screen "9" 800x480, template "Template_2"
   Button "Button_1" at 38,239 size 120x40; TextOff 'Carbamazepine'
      on Click: ActivateScreen("4_ORDER", 0); SetTag("Selected_URL", 'file:///C:/ASRS_Video/clip181.html')
      on Activate: SetTag("Selected_Medicine", 181)
      on Release: SetTag("ยา 181", 0)
      on Press: SetTag("ยา 181", 1)
   Button "Button_10" at 38,415 size 120x40; TextOff 'Pioglitazone'
      on Click: ActivateScreen("4_ORDER", 0); SetTag("Selected_URL", 'file:///C:/ASRS_Video/clip186.html')
      on Activate: SetTag("Selected_Medicine", 186)
      on Release: SetTag("ยา 186", 0)
      on Press: SetTag("ยา 186", 1)
   Button "Button_2" at 189,240 size 120x40; TextOff 'Levetiracetam'
      on Click: ActivateScreen("4_ORDER", 0); SetTag("Selected_URL", 'file:///C:/ASRS_Video/clip182.html')
      on Activate: SetTag("Selected_Medicine", 182)
      on Release: SetTag("ยา 182", 0)
      on Press: SetTag("ยา 182", 1)
   Button "Button_3" at 190,415 size 120x40; TextOff 'Sitagliptin'
      on Click: ActivateScreen("4_ORDER", 0); SetTag("Selected_URL", 'file:///C:/ASRS_Video/clip187.html')
      on Activate: SetTag("Selected_Medicine", 187)
      on Release: SetTag("ยา 187", 0)
      on Press: SetTag("ยา 187", 1)
   Button "Button_4" at 340,240 size 120x40; TextOff 'Metformin'
      on Click: ActivateScreen("4_ORDER", 0); SetTag("Selected_URL", 'file:///C:/ASRS_Video/clip183.html')
      on Activate: SetTag("Selected_Medicine", 183)
      on Release: SetTag("ยา 183", 0)
      on Press: SetTag("ยา 183", 1)
   Button "Button_5" at 340,416 size 120x40; TextOff 'Insulin regular'
      on Click: ActivateScreen("4_ORDER", 0); SetTag("Selected_URL", 'file:///C:/ASRS_Video/clip188.html')
      on Activate: SetTag("Selected_Medicine", 188)
      on Release: SetTag("ยา 188", 0)
      on Press: SetTag("ยา 188", 1)
   Button "Button_6" at 492,416 size 120x40; TextOff 'Insulin NPH'
      on Click: ActivateScreen("4_ORDER", 0); SetTag("Selected_URL", 'file:///C:/ASRS_Video/clip189.html')
      on Activate: SetTag("Selected_Medicine", 189)
      on Release: SetTag("ยา 189", 0)
      on Press: SetTag("ยา 189", 1)
   Button "Button_7" at 492,240 size 120x40; TextOff 'Glibenclamide'
      on Click: ActivateScreen("4_ORDER", 0); SetTag("Selected_URL", 'file:///C:/ASRS_Video/clip184.html')
      on Activate: SetTag("Selected_Medicine", 184)
      on Release: SetTag("ยา 184", 0)
      on Press: SetTag("ยา 184", 1)
   Button "Button_8" at 644,240 size 120x40; TextOff 'Gliclazide'
      on Click: ActivateScreen("4_ORDER", 0); SetTag("Selected_URL", 'file:///C:/ASRS_Video/clip185.html')
      on Activate: SetTag("Selected_Medicine", 185)
      on Release: SetTag("ยา 185", 0)
      on Press: SetTag("ยา 185", 1)
   Button "Button_11" at 645,416 size 120x40; TextOff 'Insulin glargine'
      on Click: ActivateScreen("4_ORDER", 0); SetTag("Selected_URL", 'file:///C:/ASRS_Video/clip190.html')
      on Activate: SetTag("Selected_Medicine", 190)
      on Release: SetTag("ยา 190", 0)
      on Press: SetTag("ยา 190", 1)
   Button "Button_12" at 24,16 size 94x40; TextOff 'Back'
      on Press: ActivateScreen("8", 0)
   Button "Button_9" at 688,16 size 96x40; TextOff 'Next'
      on Press: ActivateScreen("10", 0)
   GraphicView "Template_Graphic view_2" at 27,19 size 36x32; Picture "fast-backward"
   GraphicView "Template_Graphic view_1" at 693,20 size 36x32; Picture "play"
   GraphicView "Template_Graphic view_3" at 37,128 size 120x104; Picture "Picture181"
   GraphicView "Template_Graphic view_4" at 191,129 size 120x104; Picture "Picture182"
   GraphicView "Template_Graphic view_5" at 339,129 size 120x104; Picture "Picture183"
   GraphicView "Template_Graphic view_6" at 493,129 size 120x104; Picture "Picture184"
   GraphicView "Template_Graphic view_7" at 645,129 size 120x104; Picture "Picture185"
   GraphicView "Template_Graphic view_8" at 38,305 size 120x104; Picture "Picture186"
   GraphicView "Template_Graphic view_9" at 189,304 size 120x112; Picture "Picture187"
   GraphicView "Template_Graphic view_10" at 351,307 size 96x104; Picture "Picture188"
   GraphicView "Template_Graphic view_11" at 497,304 size 120x112; Picture "Picture189"
   GraphicView "Template_Graphic view_12" at 645,304 size 120x104; Picture "Picture190"
   TextField "Template_Text field_2" at 201,80 size 20x32; Text '9'

screen "10" 800x480, template "Template_2"
   Button "Button_1" at 38,239 size 120x40; TextOff 'Levothyroxine'
      on Click: ActivateScreen("4_ORDER", 0); SetTag("Selected_URL", 'file:///C:/ASRS_Video/clip191.html')
      on Activate: SetTag("Selected_Medicine", 191)
      on Release: SetTag("ยา 191", 0)
      on Press: SetTag("ยา 191", 1)
   Button "Button_10" at 38,415 size 120x40; TextOff 'Hydrocortisone'
      on Click: ActivateScreen("4_ORDER", 0); SetTag("Selected_URL", 'file:///C:/ASRS_Video/clip196.html')
      on Activate: SetTag("Selected_Medicine", 196)
      on Release: SetTag("ยา 196", 0)
      on Press: SetTag("ยา 196", 1)
   Button "Button_2" at 189,240 size 120x40; TextOff 'Propylthiouracil'
      on Click: ActivateScreen("4_ORDER", 0); SetTag("Selected_URL", 'file:///C:/ASRS_Video/clip192.html')
      on Activate: SetTag("Selected_Medicine", 192)
      on Release: SetTag("ยา 192", 0)
      on Press: SetTag("ยา 192", 1)
   Button "Button_3" at 190,415 size 120x40; TextOff 'Colchicine'
      on Click: ActivateScreen("4_ORDER", 0); SetTag("Selected_URL", 'file:///C:/ASRS_Video/clip197.html')
      on Activate: SetTag("Selected_Medicine", 197)
      on Release: SetTag("ยา 197", 0)
      on Press: SetTag("ยา 197", 1)
   Button "Button_4" at 340,240 size 120x40; TextOff 'Methimazole'
      on Click: ActivateScreen("4_ORDER", 0); SetTag("Selected_URL", 'file:///C:/ASRS_Video/clip193.html')
      on Activate: SetTag("Selected_Medicine", 193)
      on Release: SetTag("ยา 193", 0)
      on Press: SetTag("ยา 193", 1)
   Button "Button_5" at 340,416 size 120x40; TextOff 'Allopurinol'
      on Click: ActivateScreen("4_ORDER", 0); SetTag("Selected_URL", 'file:///C:/ASRS_Video/clip198.html')
      on Activate: SetTag("Selected_Medicine", 198)
      on Release: SetTag("ยา 198", 0)
      on Press: SetTag("ยา 198", 1)
   Button "Button_6" at 492,416 size 120x40; TextOff 'Febuxostat'
      on Click: ActivateScreen("4_ORDER", 0); SetTag("Selected_URL", 'file:///C:/ASRS_Video/clip199.html')
      on Activate: SetTag("Selected_Medicine", 199)
      on Release: SetTag("ยา 199", 0)
      on Press: SetTag("ยา 199", 1)
   Button "Button_7" at 492,240 size 120x40; TextOff 'Prednisolone'
      on Click: ActivateScreen("4_ORDER", 0); SetTag("Selected_URL", 'file:///C:/ASRS_Video/clip194.html')
      on Activate: SetTag("Selected_Medicine", 194)
      on Release: SetTag("ยา 194", 0)
      on Press: SetTag("ยา 194", 1)
   Button "Button_8" at 644,240 size 120x40; TextOff 'Dexamethasone'
      on Click: ActivateScreen("4_ORDER", 0); SetTag("Selected_URL", 'file:///C:/ASRS_Video/clip195.html')
      on Activate: SetTag("Selected_Medicine", 195)
      on Release: SetTag("ยา 195", 0)
      on Press: SetTag("ยา 195", 1)
   Button "Button_11" at 645,416 size 120x40; TextOff 'Calcium carbonate'
      on Click: ActivateScreen("4_ORDER", 0); SetTag("Selected_URL", 'file:///C:/ASRS_Video/clip200.html')
      on Activate: SetTag("Selected_Medicine", 200)
      on Release: SetTag("ยา 200", 0)
      on Press: SetTag("ยา 200", 1)
   Button "Button_12" at 24,16 size 94x40; TextOff 'Back'
      on Press: ActivateScreen("9", 0)
   Button "Button_9" at 688,16 size 96x40; TextOff 'Next'
      on Press: ActivateScreen("11", 0)
   GraphicView "Template_Graphic view_2" at 27,19 size 36x32; Picture "fast-backward"
   GraphicView "Template_Graphic view_1" at 693,20 size 36x32; Picture "play"
   GraphicView "Template_Graphic view_3" at 37,128 size 120x104; Picture "Picture191"
   GraphicView "Template_Graphic view_4" at 191,129 size 120x104; Picture "Picture192"
   GraphicView "Template_Graphic view_5" at 339,129 size 120x104; Picture "Picture193"
   GraphicView "Template_Graphic view_6" at 493,129 size 120x104; Picture "Picture194"
   GraphicView "Template_Graphic view_7" at 645,129 size 120x104; Picture "Picture195"
   GraphicView "Template_Graphic view_8" at 38,305 size 120x104; Picture "Picture196"
   GraphicView "Template_Graphic view_9" at 189,304 size 120x112; Picture "Picture197"
   GraphicView "Template_Graphic view_10" at 351,307 size 96x104; Picture "Picture198"
   GraphicView "Template_Graphic view_11" at 497,304 size 120x112; Picture "Picture199"
   GraphicView "Template_Graphic view_12" at 645,304 size 120x104; Picture "Picture200"
   TextField "Template_Text field_2" at 201,80 size 36x32; Text '10'

screen "11" 800x480, template "Template_2"
   Button "Button_1" at 38,239 size 120x40; TextOff 'Vitamin B complex'
      on Click: ActivateScreen("4_ORDER", 0); SetTag("Selected_URL", 'file:///C:/ASRS_Video/clip201.html')
      on Activate: SetTag("Selected_Medicine", 201)
      on Release: SetTag("ยา 201", 0)
      on Press: SetTag("ยา 201", 1)
   Button "Button_10" at 38,415 size 120x40; TextOff 'Potassium chloride'
      on Click: ActivateScreen("4_ORDER", 0); SetTag("Selected_URL", 'file:///C:/ASRS_Video/clip206.html')
      on Activate: SetTag("Selected_Medicine", 206)
      on Release: SetTag("ยา 206", 0)
      on Press: SetTag("ยา 206", 1)
   Button "Button_2" at 189,240 size 120x40; TextOff 'Vitamin C'
      on Click: ActivateScreen("4_ORDER", 0); SetTag("Selected_URL", 'file:///C:/ASRS_Video/clip202.html')
      on Activate: SetTag("Selected_Medicine", 202)
      on Release: SetTag("ยา 202", 0)
      on Press: SetTag("ยา 202", 1)
   Button "Button_3" at 190,415 size 120x40; TextOff 'Sodium bicarbonate'
      on Click: ActivateScreen("4_ORDER", 0); SetTag("Selected_URL", 'file:///C:/ASRS_Video/clip207.html')
      on Activate: SetTag("Selected_Medicine", 207)
      on Release: SetTag("ยา 207", 0)
      on Press: SetTag("ยา 207", 1)
   Button "Button_4" at 340,240 size 120x40; TextOff 'Ferrous fumarate'
      on Click: ActivateScreen("4_ORDER", 0); SetTag("Selected_URL", 'file:///C:/ASRS_Video/clip203.html')
      on Activate: SetTag("Selected_Medicine", 203)
      on Release: SetTag("ยา 203", 0)
      on Press: SetTag("ยา 203", 1)
   Button "Button_5" at 340,416 size 120x40; TextOff 'Calcium gluconate'
      on Click: ActivateScreen("4_ORDER", 0); SetTag("Selected_URL", 'file:///C:/ASRS_Video/clip208.html')
      on Activate: SetTag("Selected_Medicine", 208)
      on Release: SetTag("ยา 208", 0)
      on Press: SetTag("ยา 208", 1)
   Button "Button_6" at 492,416 size 120x40; TextOff 'Magnesium sulfate'
      on Click: ActivateScreen("4_ORDER", 0); SetTag("Selected_URL", 'file:///C:/ASRS_Video/clip209.html')
      on Activate: SetTag("Selected_Medicine", 209)
      on Release: SetTag("ยา 209", 0)
      on Press: SetTag("ยา 209", 1)
   Button "Button_7" at 492,240 size 120x40; TextOff 'Folic acid'
      on Click: ActivateScreen("4_ORDER", 0); SetTag("Selected_URL", 'file:///C:/ASRS_Video/clip204.html')
      on Activate: SetTag("Selected_Medicine", 204)
      on Release: SetTag("ยา 204", 0)
      on Press: SetTag("ยา 204", 1)
   Button "Button_8" at 644,240 size 120x40; TextOff 'Cyanocobalamin'
      on Click: ActivateScreen("4_ORDER", 0); SetTag("Selected_URL", 'file:///C:/ASRS_Video/clip205.html')
      on Activate: SetTag("Selected_Medicine", 205)
      on Release: SetTag("ยา 205", 0)
      on Press: SetTag("ยา 205", 1)
   Button "Button_11" at 645,416 size 120x40; TextOff 'Multivitamin'
      on Click: ActivateScreen("4_ORDER", 0); SetTag("Selected_URL", 'file:///C:/ASRS_Video/clip210.html')
      on Activate: SetTag("Selected_Medicine", 210)
      on Release: SetTag("ยา 210", 0)
      on Press: SetTag("ยา 210", 1)
   Button "Button_12" at 24,16 size 94x40; TextOff 'Back'
      on Press: ActivateScreen("10", 0)
   Button "Button_9" at 688,16 size 96x40; TextOff 'Next'
      on Press: ActivateScreen("12", 0)
   GraphicView "Template_Graphic view_2" at 27,19 size 36x32; Picture "fast-backward"
   GraphicView "Template_Graphic view_1" at 693,20 size 36x32; Picture "play"
   GraphicView "Template_Graphic view_3" at 37,128 size 120x104; Picture "Picture201"
   GraphicView "Template_Graphic view_4" at 191,129 size 120x104; Picture "Picture202"
   GraphicView "Template_Graphic view_5" at 339,129 size 120x104; Picture "Picture203"
   GraphicView "Template_Graphic view_6" at 493,129 size 120x104; Picture "Picture204"
   GraphicView "Template_Graphic view_7" at 645,129 size 120x104; Picture "Picture205"
   GraphicView "Template_Graphic view_8" at 38,305 size 120x104; Picture "Picture206"
   GraphicView "Template_Graphic view_9" at 189,304 size 120x112; Picture "Picture207"
   GraphicView "Template_Graphic view_10" at 351,307 size 96x104; Picture "Picture208"
   GraphicView "Template_Graphic view_11" at 497,304 size 120x112; Picture "Picture209"
   GraphicView "Template_Graphic view_12" at 645,304 size 120x104; Picture "Picture210"
   TextField "Template_Text field_2" at 201,80 size 36x32; Text '11'

screen "12" 800x480, template "Template_2"
   Button "Button_1" at 38,239 size 120x40; TextOff 'Oral rehydration salt'
      on Click: ActivateScreen("4_ORDER", 0); SetTag("Selected_URL", 'file:///C:/ASRS_Video/clip211.html')
      on Activate: SetTag("Selected_Medicine", 211)
      on Release: SetTag("ยา 211", 0)
      on Press: SetTag("ยา 211", 1)
   Button "Button_10" at 38,415 size 120x40; TextOff 'Piroxicam'
      on Click: ActivateScreen("4_ORDER", 0); SetTag("Selected_URL", 'file:///C:/ASRS_Video/clip216.html')
      on Activate: SetTag("Selected_Medicine", 216)
      on Release: SetTag("ยา 216", 0)
      on Press: SetTag("ยา 216", 1)
   Button "Button_2" at 189,240 size 120x40; TextOff 'Baclofen'
      on Click: ActivateScreen("4_ORDER", 0); SetTag("Selected_URL", 'file:///C:/ASRS_Video/clip212.html')
      on Activate: SetTag("Selected_Medicine", 212)
      on Release: SetTag("ยา 212", 0)
      on Press: SetTag("ยา 212", 1)
   Button "Button_3" at 190,415 size 120x40; TextOff 'Etoricoxib'
      on Click: ActivateScreen("4_ORDER", 0); SetTag("Selected_URL", 'file:///C:/ASRS_Video/clip217.html')
      on Activate: SetTag("Selected_Medicine", 217)
      on Release: SetTag("ยา 217", 0)
      on Press: SetTag("ยา 217", 1)
   Button "Button_4" at 340,240 size 120x40; TextOff 'Tizanidine'
      on Click: ActivateScreen("4_ORDER", 0); SetTag("Selected_URL", 'file:///C:/ASRS_Video/clip213.html')
      on Activate: SetTag("Selected_Medicine", 213)
      on Release: SetTag("ยา 213", 0)
      on Press: SetTag("ยา 213", 1)
   Button "Button_5" at 340,416 size 120x40; TextOff 'Glucosamine'
      on Click: ActivateScreen("4_ORDER", 0); SetTag("Selected_URL", 'file:///C:/ASRS_Video/clip218.html')
      on Activate: SetTag("Selected_Medicine", 218)
      on Release: SetTag("ยา 218", 0)
      on Press: SetTag("ยา 218", 1)
   Button "Button_6" at 492,416 size 120x40; TextOff 'Chondroitin sulfate'
      on Click: ActivateScreen("4_ORDER", 0); SetTag("Selected_URL", 'file:///C:/ASRS_Video/clip219.html')
      on Activate: SetTag("Selected_Medicine", 219)
      on Release: SetTag("ยา 219", 0)
      on Press: SetTag("ยา 219", 1)
   Button "Button_7" at 492,240 size 120x40; TextOff 'Orphenadrine'
      on Click: ActivateScreen("4_ORDER", 0); SetTag("Selected_URL", 'file:///C:/ASRS_Video/clip214.html')
      on Activate: SetTag("Selected_Medicine", 214)
      on Release: SetTag("ยา 214", 0)
      on Press: SetTag("ยา 214", 1)
   Button "Button_8" at 644,240 size 120x40; TextOff 'Meloxicam'
      on Click: ActivateScreen("4_ORDER", 0); SetTag("Selected_URL", 'file:///C:/ASRS_Video/clip215.html')
      on Activate: SetTag("Selected_Medicine", 215)
      on Release: SetTag("ยา 215", 0)
      on Press: SetTag("ยา 215", 1)
   Button "Button_11" at 645,416 size 120x40; TextOff 'Alendronate'
      on Click: ActivateScreen("4_ORDER", 0); SetTag("Selected_URL", 'file:///C:/ASRS_Video/clip220.html')
      on Activate: SetTag("Selected_Medicine", 220)
      on Release: SetTag("ยา 220", 0)
      on Press: SetTag("ยา 220", 1)
   Button "Button_12" at 24,16 size 94x40; TextOff 'Back'
      on Press: ActivateScreen("11", 0)
   GraphicView "Template_Graphic view_2" at 27,19 size 36x32; Picture "fast-backward"
   GraphicView "Template_Graphic view_3" at 37,128 size 120x104; Picture "Picture211"
   GraphicView "Template_Graphic view_4" at 191,129 size 120x104; Picture "Picture212"
   GraphicView "Template_Graphic view_5" at 339,129 size 120x104; Picture "Picture213"
   GraphicView "Template_Graphic view_6" at 493,129 size 120x104; Picture "Picture214"
   GraphicView "Template_Graphic view_7" at 645,129 size 120x104; Picture "Picture215"
   GraphicView "Template_Graphic view_8" at 38,305 size 120x104; Picture "Picture216"
   GraphicView "Template_Graphic view_9" at 189,304 size 120x112; Picture "Picture217"
   GraphicView "Template_Graphic view_10" at 351,307 size 96x104; Picture "Picture218"
   GraphicView "Template_Graphic view_11" at 497,304 size 120x112; Picture "Picture219"
   GraphicView "Template_Graphic view_12" at 645,304 size 120x104; Picture "Picture220"
   TextField "Template_Text field_2" at 201,80 size 36x32; Text '12'

screen "1_3" 800x480, template "Template_2"
   Button "Button_1" at 40,240 size 120x40; TextOff 'Artificial tears'
      on Click: ActivateScreen("4_ORDER", 0); SetTag("Selected_URL", 'file:///C:/ASRS_Video/clip461.html')
      on Activate: SetTag("Selected_Medicine", 461)
      on Release: SetTag("ยา 461", 0)
      on Press: SetTag("ยา 461", 1)
   Button "Button_10" at 38,415 size 120x40; TextOff 'Timolol'
      on Click: ActivateScreen("4_ORDER", 0); SetTag("Selected_URL", 'file:///C:/ASRS_Video/clip466.html')
      on Activate: SetTag("Selected_Medicine", 466)
      on Release: SetTag("ยา 466", 0)
      on Press: SetTag("ยา 466", 1)
   Button "Button_2" at 189,240 size 120x40; TextOff 'Carboxy methylcellulose'
      on Click: ActivateScreen("4_ORDER", 0); SetTag("Selected_URL", 'file:///C:/ASRS_Video/clip462.html')
      on Activate: SetTag("Selected_Medicine", 462)
      on Release: SetTag("ยา 462", 0)
      on Press: SetTag("ยา 462", 1)
   Button "Button_3" at 190,415 size 120x40; TextOff 'Betaxolol'
      on Click: ActivateScreen("4_ORDER", 0); SetTag("Selected_URL", 'file:///C:/ASRS_Video/clip467.html')
      on Activate: SetTag("Selected_Medicine", 467)
      on Release: SetTag("ยา 467", 0)
      on Press: SetTag("ยา 467", 1)
   Button "Button_4" at 340,240 size 120x40; TextOff 'Hydroxypropyl methylcellulose'
      on Click: ActivateScreen("4_ORDER", 0); SetTag("Selected_URL", 'file:///C:/ASRS_Video/clip463.html')
      on Activate: SetTag("Selected_Medicine", 463)
      on Release: SetTag("ยา 463", 0)
      on Press: SetTag("ยา 463", 1)
   Button "Button_5" at 340,416 size 120x40; TextOff 'Brimonidine'
      on Click: ActivateScreen("4_ORDER", 0); SetTag("Selected_URL", 'file:///C:/ASRS_Video/clip468.html')
      on Activate: SetTag("Selected_Medicine", 468)
      on Release: SetTag("ยา 468", 0)
      on Press: SetTag("ยา 468", 1)
   Button "Button_6" at 492,416 size 120x40; TextOff 'Dorzolamide'
      on Click: ActivateScreen("4_ORDER", 0); SetTag("Selected_URL", 'file:///C:/ASRS_Video/clip469.html')
      on Activate: SetTag("Selected_Medicine", 469)
      on Release: SetTag("ยา 469", 0)
      on Press: SetTag("ยา 469", 1)
   Button "Button_7" at 492,240 size 120x40; TextOff 'Sodium hyaluronate'
      on Click: ActivateScreen("4_ORDER", 0); SetTag("Selected_URL", 'file:///C:/ASRS_Video/clip464.html')
      on Activate: SetTag("Selected_Medicine", 464)
      on Release: SetTag("ยา 464", 0)
      on Press: SetTag("ยา 464", 1)
   Button "Button_8" at 644,240 size 120x40; TextOff 'Polyvinyl alcohol'
      on Click: ActivateScreen("4_ORDER", 0); SetTag("Selected_URL", 'file:///C:/ASRS_Video/clip465.html')
      on Activate: SetTag("Selected_Medicine", 465)
      on Release: SetTag("ยา 465", 0)
      on Press: SetTag("ยา 465", 1)
   Button "Button_11" at 645,416 size 120x40; TextOff 'Acetazolamide'
      on Click: ActivateScreen("4_ORDER", 0); SetTag("Selected_URL", 'file:///C:/ASRS_Video/clip470.html')
      on Activate: SetTag("Selected_Medicine", 470)
      on Release: SetTag("ยา 470", 0)
      on Press: SetTag("ยา 470", 1)
   Button "Button_12" at 688,16 size 96x40; TextOff 'Next'
      on Press: ActivateScreen("2_3", 0)
   Button "Button_9" at 24,16 size 94x40; TextOff 'Back'
      on Press: ActivateScreen("4_ORDER", 0)
   GraphicView "Template_Graphic view_2" at 693,20 size 36x32; Picture "play"
   GraphicView "Template_Graphic view_1" at 27,19 size 36x32; Picture "fast-backward"
   GraphicView "Template_Graphic view_3" at 37,128 size 120x104; Picture "1_2"
   GraphicView "Template_Graphic view_4" at 191,129 size 120x104; Picture "2_2"
   GraphicView "Template_Graphic view_5" at 339,129 size 120x104; Picture "3_2"
   GraphicView "Template_Graphic view_6" at 493,129 size 120x104; Picture "4_2"
   GraphicView "Template_Graphic view_7" at 645,129 size 120x104; Picture "5_2"
   GraphicView "Template_Graphic view_8" at 38,305 size 120x104; Picture "6_2"
   GraphicView "Template_Graphic view_9" at 189,304 size 120x112; Picture "7_2"
   GraphicView "Template_Graphic view_10" at 351,307 size 96x104; Picture "8_2"
   GraphicView "Template_Graphic view_11" at 497,304 size 120x112; Picture "9_2"
   GraphicView "Template_Graphic view_12" at 645,304 size 120x104; Picture "10_2"
   TextField "Template_Text field_2" at 201,80 size 20x32; Text '1'

screen "2_3" 800x480, template "Template_2"
   Button "Button_1" at 38,239 size 120x40; TextOff 'Latanoprost'
      on Click: ActivateScreen("4_ORDER", 0); SetTag("Selected_URL", 'file:///C:/ASRS_Video/clip471.html')
      on Activate: SetTag("Selected_Medicine", 471)
      on Release: SetTag("ยา 471", 0)
      on Press: SetTag("ยา 471", 1)
   Button "Button_9" at 688,16 size 96x40; TextOff 'Next'
      on Press: ActivateScreen("3_3", 0)
   Button "Button_10" at 38,415 size 120x40; TextOff 'Tropicamide'
      on Click: ActivateScreen("4_ORDER", 0); SetTag("Selected_URL", 'file:///C:/ASRS_Video/clip476.html')
      on Activate: SetTag("Selected_Medicine", 476)
      on Release: SetTag("ยา 476", 0)
      on Press: SetTag("ยา 476", 1)
   Button "Button_2" at 189,240 size 120x40; TextOff 'Travoprost'
      on Click: ActivateScreen("4_ORDER", 0); SetTag("Selected_URL", 'file:///C:/ASRS_Video/clip472.html')
      on Activate: SetTag("Selected_Medicine", 472)
      on Release: SetTag("ยา 472", 0)
      on Press: SetTag("ยา 472", 1)
   Button "Button_3" at 190,415 size 120x40; TextOff 'Phenylephrine'
      on Click: ActivateScreen("4_ORDER", 0); SetTag("Selected_URL", 'file:///C:/ASRS_Video/clip477.html')
      on Activate: SetTag("Selected_Medicine", 477)
      on Release: SetTag("ยา 477", 0)
      on Press: SetTag("ยา 477", 1)
   Button "Button_4" at 340,240 size 120x40; TextOff 'Bimatoprost'
      on Click: ActivateScreen("4_ORDER", 0); SetTag("Selected_URL", 'file:///C:/ASRS_Video/clip473.html')
      on Activate: SetTag("Selected_Medicine", 473)
      on Release: SetTag("ยา 473", 0)
      on Press: SetTag("ยา 473", 1)
   Button "Button_5" at 340,416 size 120x40; TextOff 'Ciprofloxacin'
      on Click: ActivateScreen("4_ORDER", 0); SetTag("Selected_URL", 'file:///C:/ASRS_Video/clip478.html')
      on Activate: SetTag("Selected_Medicine", 478)
      on Release: SetTag("ยา 478", 0)
      on Press: SetTag("ยา 478", 1)
   Button "Button_6" at 492,416 size 120x40; TextOff 'Ofloxacin'
      on Click: ActivateScreen("4_ORDER", 0); SetTag("Selected_URL", 'file:///C:/ASRS_Video/clip479.html')
      on Activate: SetTag("Selected_Medicine", 479)
      on Release: SetTag("ยา 479", 0)
      on Press: SetTag("ยา 479", 1)
   Button "Button_7" at 492,240 size 120x40; TextOff 'Pilocarpine'
      on Click: ActivateScreen("4_ORDER", 0); SetTag("Selected_URL", 'file:///C:/ASRS_Video/clip474.html')
      on Activate: SetTag("Selected_Medicine", 474)
      on Release: SetTag("ยา 474", 0)
      on Press: SetTag("ยา 474", 1)
   Button "Button_8" at 644,240 size 120x40; TextOff 'Atropine'
      on Click: ActivateScreen("4_ORDER", 0); SetTag("Selected_URL", 'file:///C:/ASRS_Video/clip475.html')
      on Activate: SetTag("Selected_Medicine", 475)
      on Release: SetTag("ยา 475", 0)
      on Press: SetTag("ยา 475", 1)
   Button "Button_11" at 645,416 size 120x40; TextOff 'Moxifloxacin'
      on Click: ActivateScreen("4_ORDER", 0); SetTag("Selected_URL", 'file:///C:/ASRS_Video/clip480.html')
      on Activate: SetTag("Selected_Medicine", 480)
      on Release: SetTag("ยา 480", 0)
      on Press: SetTag("ยา 480", 1)
   Button "Button_12" at 24,16 size 94x40; TextOff 'Back'
      on Press: ActivateScreen("1_3", 0)
   GraphicView "Template_Graphic view_1" at 693,20 size 36x32; Picture "play"
   GraphicView "Template_Graphic view_2" at 27,19 size 36x32; Picture "fast-backward"
   GraphicView "Template_Graphic view_3" at 37,128 size 120x104; Picture "11_2"
   GraphicView "Template_Graphic view_4" at 191,129 size 120x104; Picture "12_2"
   GraphicView "Template_Graphic view_5" at 339,129 size 120x104; Picture "13_2"
   GraphicView "Template_Graphic view_6" at 493,129 size 120x104; Picture "14_2"
   GraphicView "Template_Graphic view_7" at 645,129 size 120x104; Picture "15_2"
   GraphicView "Template_Graphic view_8" at 38,305 size 120x104; Picture "16_2"
   GraphicView "Template_Graphic view_9" at 189,304 size 120x112; Picture "17_2"
   GraphicView "Template_Graphic view_10" at 351,307 size 96x104; Picture "18_2"
   GraphicView "Template_Graphic view_11" at 497,304 size 120x112; Picture "19_2"
   GraphicView "Template_Graphic view_12" at 645,304 size 120x104; Picture "20_2"
   TextField "Template_Text field_2" at 201,80 size 20x32; Text '2'

screen "3_3" 800x480, template "Template_2"
   Button "Button_1" at 38,239 size 120x40; TextOff 'Tobramycin'
      on Click: ActivateScreen("4_ORDER", 0); SetTag("Selected_URL", 'file:///C:/ASRS_Video/clip481.html')
      on Activate: SetTag("Selected_Medicine", 481)
      on Release: SetTag("ยา 481", 0)
      on Press: SetTag("ยา 481", 1)
   Button "Button_9" at 688,16 size 96x40; TextOff 'Next'
      on Press: ActivateScreen("4_3", 0)
   Button "Button_10" at 38,415 size 120x40; TextOff 'Acyclovir'
      on Click: ActivateScreen("4_ORDER", 0); SetTag("Selected_URL", 'file:///C:/ASRS_Video/clip486.html')
      on Activate: SetTag("Selected_Medicine", 486)
      on Release: SetTag("ยา 486", 0)
      on Press: SetTag("ยา 486", 1)
   Button "Button_2" at 189,240 size 120x40; TextOff 'Gentamicin'
      on Click: ActivateScreen("4_ORDER", 0); SetTag("Selected_URL", 'file:///C:/ASRS_Video/clip482.html')
      on Activate: SetTag("Selected_Medicine", 482)
      on Release: SetTag("ยา 482", 0)
      on Press: SetTag("ยา 482", 1)
   Button "Button_3" at 190,415 size 120x40; TextOff 'Prednisolone acetate'
      on Click: ActivateScreen("4_ORDER", 0); SetTag("Selected_URL", 'file:///C:/ASRS_Video/clip487.html')
      on Activate: SetTag("Selected_Medicine", 487)
      on Release: SetTag("ยา 487", 0)
      on Press: SetTag("ยา 487", 1)
   Button "Button_4" at 340,240 size 120x40; TextOff 'Chloramphenicol'
      on Click: ActivateScreen("4_ORDER", 0); SetTag("Selected_URL", 'file:///C:/ASRS_Video/clip483.html')
      on Activate: SetTag("Selected_Medicine", 483)
      on Release: SetTag("ยา 483", 0)
      on Press: SetTag("ยา 483", 1)
   Button "Button_5" at 340,416 size 120x40; TextOff 'Dexamethasone'
      on Click: ActivateScreen("4_ORDER", 0); SetTag("Selected_URL", 'file:///C:/ASRS_Video/clip488.html')
      on Activate: SetTag("Selected_Medicine", 488)
      on Release: SetTag("ยา 488", 0)
      on Press: SetTag("ยา 488", 1)
   Button "Button_6" at 492,416 size 120x40; TextOff 'Fluorometholone'
      on Click: ActivateScreen("4_ORDER", 0); SetTag("Selected_URL", 'file:///C:/ASRS_Video/clip489.html')
      on Activate: SetTag("Selected_Medicine", 489)
      on Release: SetTag("ยา 489", 0)
      on Press: SetTag("ยา 489", 1)
   Button "Button_7" at 492,240 size 120x40; TextOff 'Fusidic acid'
      on Click: ActivateScreen("4_ORDER", 0); SetTag("Selected_URL", 'file:///C:/ASRS_Video/clip484.html')
      on Activate: SetTag("Selected_Medicine", 484)
      on Release: SetTag("ยา 484", 0)
      on Press: SetTag("ยา 484", 1)
   Button "Button_8" at 644,240 size 120x40; TextOff 'Natamycin'
      on Click: ActivateScreen("4_ORDER", 0); SetTag("Selected_URL", 'file:///C:/ASRS_Video/clip485.html')
      on Activate: SetTag("Selected_Medicine", 485)
      on Release: SetTag("ยา 485", 0)
      on Press: SetTag("ยา 485", 1)
   Button "Button_11" at 645,416 size 120x40; TextOff 'Ketorolac'
      on Click: ActivateScreen("4_ORDER", 0); SetTag("Selected_URL", 'file:///C:/ASRS_Video/clip490.html')
      on Activate: SetTag("Selected_Medicine", 490)
      on Release: SetTag("ยา 490", 0)
      on Press: SetTag("ยา 490", 1)
   Button "Button_12" at 24,16 size 94x40; TextOff 'Back'
      on Press: ActivateScreen("2_3", 0)
   GraphicView "Template_Graphic view_1" at 693,20 size 36x32; Picture "play"
   GraphicView "Template_Graphic view_2" at 27,19 size 36x32; Picture "fast-backward"
   GraphicView "Template_Graphic view_3" at 37,128 size 120x104; Picture "21_2"
   GraphicView "Template_Graphic view_4" at 191,129 size 120x104; Picture "22_2"
   GraphicView "Template_Graphic view_5" at 339,129 size 120x104; Picture "23_2"
   GraphicView "Template_Graphic view_6" at 493,129 size 120x104; Picture "24_2"
   GraphicView "Template_Graphic view_7" at 645,129 size 120x104; Picture "25_2"
   GraphicView "Template_Graphic view_8" at 38,305 size 120x104; Picture "26_2"
   GraphicView "Template_Graphic view_9" at 189,304 size 120x112; Picture "27_2"
   GraphicView "Template_Graphic view_10" at 351,307 size 96x104; Picture "28_2"
   GraphicView "Template_Graphic view_11" at 497,304 size 120x112; Picture "29_2"
   GraphicView "Template_Graphic view_12" at 645,304 size 120x104; Picture "30_2"
   TextField "Template_Text field_2" at 201,80 size 20x32; Text '3'

screen "4_3" 800x480, template "Template_2"
   Button "Button_1" at 38,239 size 120x40; TextOff 'Diclofenac'
      on Click: ActivateScreen("4_ORDER", 0); SetTag("Selected_URL", 'file:///C:/ASRS_Video/clip491.html')
      on Activate: SetTag("Selected_Medicine", 491)
      on Release: SetTag("ยา 491", 0)
      on Press: SetTag("ยา 491", 1)
   Button "Button_2" at 189,240 size 120x40; TextOff 'Olopatadine'
      on Click: ActivateScreen("4_ORDER", 0); SetTag("Selected_URL", 'file:///C:/ASRS_Video/clip492.html')
      on Activate: SetTag("Selected_Medicine", 492)
      on Release: SetTag("ยา 492", 0)
      on Press: SetTag("ยา 492", 1)
   Button "Button_4" at 340,240 size 120x40; TextOff 'Ketotifen'
      on Click: ActivateScreen("4_ORDER", 0); SetTag("Selected_URL", 'file:///C:/ASRS_Video/clip493.html')
      on Activate: SetTag("Selected_Medicine", 493)
      on Release: SetTag("ยา 493", 0)
      on Press: SetTag("ยา 493", 1)
   Button "Button_7" at 492,240 size 120x40; TextOff 'Sodium cromoglycate'
      on Click: ActivateScreen("4_ORDER", 0); SetTag("Selected_URL", 'file:///C:/ASRS_Video/clip494.html')
      on Activate: SetTag("Selected_Medicine", 494)
      on Release: SetTag("ยา 494", 0)
      on Press: SetTag("ยา 494", 1)
   Button "Button_12" at 24,16 size 94x40; TextOff 'Back'
      on Press: ActivateScreen("3_3", 0)
   GraphicView "Template_Graphic view_2" at 27,19 size 36x32; Picture "fast-backward"
   GraphicView "Template_Graphic view_3" at 37,128 size 120x104; Picture "31_2"
   GraphicView "Template_Graphic view_4" at 191,129 size 120x104; Picture "32_2"
   GraphicView "Template_Graphic view_5" at 339,129 size 120x104; Picture "33_2"
   GraphicView "Template_Graphic view_6" at 493,129 size 120x104; Picture "34_2"
   TextField "Template_Text field_2" at 201,80 size 20x32; Text '4'

screen "5_3" 800x480, template "Template_2"
   Button "Button_1" at 38,239 size 120x40; TextOff 'Mometasone'
      on Click: ActivateScreen("4_ORDER", 0)
      on Activate: SetTag("Selected_Medicine", 501)
      on Release: SetTag("ยา 501", 0)
      on Press: SetTag("ยา 501", 1)
   Button "Button_9" at 688,16 size 96x40; TextOff 'Next'
      on Press: ActivateScreen("6_3", 0)
   Button "Button_10" at 38,415 size 120x40; TextOff 'Menthol inhaler'
      on Click: ActivateScreen("4_ORDER", 0)
      on Activate: SetTag("Selected_Medicine", 506)
      on Release: SetTag("ยา 506", 0)
      on Press: SetTag("ยา 506", 1)
   Button "Button_2" at 189,240 size 120x40; TextOff 'Budesonide'
      on Click: ActivateScreen("4_ORDER", 0)
      on Activate: SetTag("Selected_Medicine", 502)
      on Release: SetTag("ยา 502", 0)
      on Press: SetTag("ยา 502", 1)
   Button "Button_3" at 190,415 size 120x40; TextOff 'Carbamide peroxide'
      on Click: ActivateScreen("4_ORDER", 0)
      on Activate: SetTag("Selected_Medicine", 507)
      on Release: SetTag("ยา 507", 0)
      on Press: SetTag("ยา 507", 1)
   Button "Button_4" at 340,240 size 120x40; TextOff 'Beclomethasone'
      on Click: ActivateScreen("4_ORDER", 0)
      on Activate: SetTag("Selected_Medicine", 503)
      on Release: SetTag("ยา 503", 0)
      on Press: SetTag("ยา 503", 1)
   Button "Button_5" at 340,416 size 120x40; TextOff 'Brinzolamide'
      on Click: ActivateScreen("4_ORDER", 0)
      on Activate: SetTag("Selected_Medicine", 508)
      on Release: SetTag("ยา 508", 0)
      on Press: SetTag("ยา 508", 1)
   Button "Button_6" at 492,416 size 120x40; TextOff 'Ciprofloxacin'
      on Click: ActivateScreen("4_ORDER", 0)
      on Activate: SetTag("Selected_Medicine", 509)
      on Release: SetTag("ยา 509", 0)
      on Press: SetTag("ยา 509", 1)
   Button "Button_7" at 492,240 size 120x40; TextOff 'Azelastine'
      on Click: ActivateScreen("4_ORDER", 0)
      on Activate: SetTag("Selected_Medicine", 504)
      on Release: SetTag("ยา 504", 0)
      on Press: SetTag("ยา 504", 1)
   Button "Button_8" at 644,240 size 120x40; TextOff 'Ipratropium bromide'
      on Click: ActivateScreen("4_ORDER", 0)
      on Activate: SetTag("Selected_Medicine", 505)
      on Release: SetTag("ยา 505", 0)
      on Press: SetTag("ยา 505", 1)
   Button "Button_11" at 645,416 size 120x40; TextOff 'Ofloxacin'
      on Click: ActivateScreen("4_ORDER", 0)
      on Activate: SetTag("Selected_Medicine", 510)
      on Release: SetTag("ยา 510", 0)
      on Press: SetTag("ยา 510", 1)
   Button "Button_12" at 24,16 size 94x40; TextOff 'Back'
      on Press: ActivateScreen("4_3", 0)
   GraphicView "Template_Graphic view_1" at 693,20 size 36x32; Picture "play"
   GraphicView "Template_Graphic view_2" at 27,19 size 36x32; Picture "fast-backward"
   GraphicView "Template_Graphic view_3" at 37,128 size 120x104; Picture "41_2"
   GraphicView "Template_Graphic view_4" at 191,129 size 120x104; Picture "42_2"
   GraphicView "Template_Graphic view_5" at 339,129 size 120x104; Picture "43_2"
   GraphicView "Template_Graphic view_6" at 493,129 size 120x104; Picture "44_2"
   GraphicView "Template_Graphic view_7" at 645,129 size 120x104; Picture "45_2"
   GraphicView "Template_Graphic view_8" at 38,305 size 120x104; Picture "46_2"
   GraphicView "Template_Graphic view_9" at 189,304 size 120x112; Picture "47_2"
   GraphicView "Template_Graphic view_10" at 351,307 size 96x104; Picture "48_2"
   GraphicView "Template_Graphic view_11" at 497,304 size 120x112; Picture "49_2"
   GraphicView "Template_Graphic view_12" at 645,304 size 120x104; Picture "50_2"
   TextField "Template_Text field_2" at 201,80 size 20x32; Text '5'

screen "6_3" 800x480, template "Template_2"
   Button "Button_1" at 38,239 size 120x40; TextOff 'Neomycin polymyxin hydrocortisone'
      on Click: ActivateScreen("4_ORDER", 0)
      on Activate: SetTag("Selected_Medicine", 511)
      on Release: SetTag("ยา 511", 0)
      on Press: SetTag("ยา 511", 1)
   Button "Button_10" at 38,415 size 120x40; TextOff 'Nystatin'
      on Click: ActivateScreen("4_ORDER", 0)
      on Activate: SetTag("Selected_Medicine", 516)
      on Release: SetTag("ยา 516", 0)
      on Press: SetTag("ยา 516", 1)
   Button "Button_2" at 189,240 size 120x40; TextOff 'Lidocaine'
      on Click: ActivateScreen("4_ORDER", 0)
      on Activate: SetTag("Selected_Medicine", 512)
      on Release: SetTag("ยา 512", 0)
      on Press: SetTag("ยา 512", 1)
   Button "Button_3" at 190,415 size 120x40; TextOff 'Miconazole'
      on Click: ActivateScreen("4_ORDER", 0)
      on Activate: SetTag("Selected_Medicine", 517)
      on Release: SetTag("ยา 517", 0)
      on Press: SetTag("ยา 517", 1)
   Button "Button_4" at 340,240 size 120x40; TextOff 'Benzydamine'
      on Click: ActivateScreen("4_ORDER", 0)
      on Activate: SetTag("Selected_Medicine", 513)
      on Release: SetTag("ยา 513", 0)
      on Press: SetTag("ยา 513", 1)
   Button "Button_5" at 340,416 size 120x40; TextOff 'Triamcinolone acetonide'
      on Click: ActivateScreen("4_ORDER", 0)
      on Activate: SetTag("Selected_Medicine", 518)
      on Release: SetTag("ยา 518", 0)
      on Press: SetTag("ยา 518", 1)
   Button "Button_6" at 492,416 size 120x40; TextOff 'Lidocaine viscous'
      on Click: ActivateScreen("4_ORDER", 0)
      on Activate: SetTag("Selected_Medicine", 519)
      on Release: SetTag("ยา 519", 0)
      on Press: SetTag("ยา 519", 1)
   Button "Button_7" at 492,240 size 120x40; TextOff 'Chlorhexidine'
      on Click: ActivateScreen("4_ORDER", 0)
      on Activate: SetTag("Selected_Medicine", 514)
      on Release: SetTag("ยา 514", 0)
      on Press: SetTag("ยา 514", 1)
   Button "Button_8" at 644,240 size 120x40; TextOff 'Povidone iodine'
      on Click: ActivateScreen("4_ORDER", 0)
      on Activate: SetTag("Selected_Medicine", 515)
      on Release: SetTag("ยา 515", 0)
      on Press: SetTag("ยา 515", 1)
   Button "Button_11" at 645,416 size 120x40; TextOff 'Sodium fluoride'
      on Click: ActivateScreen("4_ORDER", 0)
      on Activate: SetTag("Selected_Medicine", 520)
      on Release: SetTag("ยา 520", 0)
      on Press: SetTag("ยา 520", 1)
   Button "Button_12" at 24,16 size 94x40; TextOff 'Back'
      on Press: ActivateScreen("5_3", 0)
   GraphicView "Template_Graphic view_2" at 27,19 size 36x32; Picture "fast-backward"
   GraphicView "Template_Graphic view_3" at 37,128 size 120x104; Picture "51_2"
   GraphicView "Template_Graphic view_4" at 191,129 size 120x104; Picture "52_2"
   GraphicView "Template_Graphic view_5" at 339,129 size 120x104; Picture "53_2"
   GraphicView "Template_Graphic view_6" at 493,129 size 120x104; Picture "54_2"
   GraphicView "Template_Graphic view_7" at 645,129 size 120x104; Picture "55_2"
   GraphicView "Template_Graphic view_8" at 38,305 size 120x104; Picture "56_2"
   GraphicView "Template_Graphic view_9" at 189,304 size 120x112; Picture "57_2"
   GraphicView "Template_Graphic view_10" at 351,307 size 96x104; Picture "58_2"
   GraphicView "Template_Graphic view_11" at 497,304 size 120x112; Picture "59_2"
   GraphicView "Template_Graphic view_12" at 645,304 size 120x104; Picture "60_2"
   TextField "Template_Text field_2" at 201,80 size 20x32; Text '6'

screen "4_ORDER" 800x480, template "ORDER"
   SymbolicIOField "Symbolic I/O field_1" at 376,204 size 386x72; TextOn '1'; TextOff '0'; TextList "SelectedMedicine"
      ProcessValue <- "แสดงชื่อยา"
   Button "Button_4" at 16,64 size 320x64; TextOn 'ยาแก้ปวด / ลดไข้'; TextOff 'ยาสำหรับหัตถการและฉุกเฉิน (Procedural & Emergency)'
      on Press: ActivateScreen("1-10", 0)
   Button "Button_5" at 16,131 size 320x64; TextOn 'ยาทาภายนอก / ผิวหนัง'; TextOff 'ยาต้านการติดเชื้อและวัคซีน (Anti-infective Immunological)'
      on Press: ActivateScreen("1_1", 0)
   Button "Button_6" at 17,198 size 320x64; TextOn 'วิตามิน / อาหารเสริม'; TextOff 'ยาเฉพาะทางและมะเร็ง (Specialized & Oncology)'
      on Press: ActivateScreen("1_2", 0)
   Button "Button_7" at 18,265 size 320x64; TextOn 'กลุ่มยาระบบทางเดินอาหาร'; TextOff 'ยารักษาโรคทั่วไป (General Medicine)'
      on Press: ActivateScreen("1", 0)
   Button "Button_3" at 16,405 size 120x68; TextOff 'HOME'
      on Press: ActivateScreen("1_OVERVIEW_1", 0)
   Button "Button_1" at 144,405 size 192x68; TextOff 'Status System'
      on Click: ActivateScreen("Status System", 0)
   Button "Button_2" at 19,332 size 320x64; TextOn 'กลุ่มยาระบบทางเดินอาหาร'; TextOff 'ยาใช้ภายนอกและอวัยวะเฉพาะ (Topical & Sensory Organ)'
      on Press: ActivateScreen("1_3", 0)
   GraphicView "Template_Graphic view_1" at 21,68 size 63x56; Picture "Med"
   GraphicView "Template_Graphic view_2" at 24,136 size 55x48; Picture "tube"
   GraphicView "Template_Graphic view_3" at 25,202 size 63x56; Picture "vitamins"
   GraphicView "Template_Graphic view_4" at 23,269 size 63x56; Picture "medicine-pills"
   Button "Template_Button_3" at 368,368 size 192x88; TextOff 'CLEAR'
      on Release: SetTag("ปุ่มClear", 0)
      on Press: SetTag("ปุ่มClear", 1)
   Button "Template_Button_1" at 568,368 size 192x88; TextOff 'CONFIRM'
      on Click: function_efd93a16("Confirm", 0, 0, 1, -1, 1); ActivateScreen("Status System", 0)
      on Press: SetTag("ปุ่มยืนยันหน้า Screen", 1)
      on Release: SetTag("ปุ่มยืนยันหน้า Screen", 0)
      on Activate: "Retrieval"()
   GraphicView "Template_Graphic view_5" at 20,416 size 46x41; Picture "NEW_HOME"
   GraphicView "Template_Graphic view_6" at 156,416 size 46x41; Picture "development"
   GraphicView "Template_Graphic view_7" at 27,336 size 63x56; Picture "drugs"

screen "2_ALAREMS" 800x480, template "Alarms"
   AlarmView "Alarm view_1" at 24,96 size 744x308
   Button "Back" at 19,409 size 159x47; TextOn 'Back'; TextOff 'Back'
      on Press: ActivateScreen("Status System", 0)
   Button "Back_1" at 612,408 size 159x47; TextOn 'Back'; TextOff 'Home'
      on Press: ActivateScreen("1_OVERVIEW_1", 0)

screen "1_OVERVIEW_1" 800x480, template "Template"
   Button "Button_3" at 668,146 size 128x48; TextOff 'STOCK'
      on Press: ActivateScreen("Screen_1", 0)
   Button "Button_4" at 668,196 size 128x48; TextOff 'RET'
      on Press: ActivateScreen("4_ORDER", 0)
   Button "Button_5" at 668,246 size 128x48; TextOff 'property'
      on Press: ActivateScreen(" propertyเบิกจ่าย", 0)
   Button "Button_6" at 668,296 size 128x48; TextOn 'LOGOUT'; TextOff 'LOGOUT'
      on Activate: function_f23ef4c9(); ActivateScreen("LOGIN", 0)
   Button "Button_1" at 668,96 size 128x48; TextOff 'Status System'
      on Click: ActivateScreen("Status System", 0)
   Button "Button_7" at 668,346 size 128x32; TextOn 'RESET'; TextOff 'Text'
      on Press: SetTag("Reset-All System", 1)
      on Release: SetTag("Reset-All System", 0)
   GraphicView "Template_Graphic view_2" at 677,153 size 35x32; Picture "management"
   GraphicView "Template_Graphic view_3" at 672,198 size 52x48; Picture "Med"
   GraphicView "Template_Graphic view_4" at 680,254 size 36x32; Picture "st"
   GraphicView "Template_Graphic view_5" at 675,300 size 45x40; Picture "logout"
   GraphicView "Template_Graphic view_6" at 675,104 size 38x33; Picture "development"
   GraphicView "Template_Graphic view_1" at 686,387 size 93x87; Picture "emergency"
   TextField "Text field_1" at 712,352 size 47x18; Text 'RESET'
   Button "Button_2" at 680,386 size 104x88; TextOff 'Text'
      on Click: InvertBit("Emergency stop")

screen " propertyจัดเก็บ" 800x480, template "property HMI data"
   SymbolicIOField "Template_Symbolic I/O field_2" at 19,249 size 122x32; TextOn '1'; TextOff '0'; TextList "X AXIS ( Horizontall )จัดเก็บ"
      ProcessValue <- "แสดงชื่อยา2"
   SymbolicIOField "Template_Symbolic I/O field_3" at 18,380 size 122x32; TextOn '1'; TextOff '0'; TextList "Y AXIS ( Verticall )จัดเก็บ"
      ProcessValue <- "แสดงชื่อยา2"
   Circle "Template_Circle_5" at 104,87 size 56x56
      Appearance <- "ป้อนรหัส Barcode"
   Circle "Template_Circle_2" at 177,88 size 56x56
      Appearance <- "Gripperเคลื่อนที่มาเอายา"
   Circle "Template_Circle_4" at 248,88 size 56x56
      Appearance <- "Gripper เคลื่อนไปช่องยา"
   Circle "Template_Circle_7" at 320,87 size 56x56
      Appearance <- "Gripper วางยา"
   Button "Template_Button_2" at 672,89 size 112x64; TextOff 'Medicine Retrieval'
      on Click: ActivateScreen(" propertyเบิกจ่าย", 0)
   SymbolicIOField "Template_Symbolic I/O field_23" at 97,293 size 74x24; TextOn '1'; TextOff '0'; TextList "EncoderแกนX (จัดเก็บ)"
      ProcessValue <- "แสดงชื่อยา2"
   SymbolicIOField "Template_Symbolic I/O field_24" at 98,428 size 74x24; TextOn '1'; TextOff '0'; TextList "EncoderแกนY (จัดเก็บ)"
      ProcessValue <- "แสดงชื่อยา2"
   Button "Template_Button_3" at 560,368 size 112x24; TextOff 'Reset to Default'
   Button "Template_Button_4" at 560,408 size 112x24; TextOff 'MODIFY'
   Button "Template_Button_1" at 681,422 size 88x24; TextOff 'HOME'
      on Press: ActivateScreen("1_OVERVIEW_1", 0)
   Button "Template_Button_5" at 681,358 size 88x24; TextOff 'START'
   Button "Template_Button_6" at 681,388 size 88x24; TextOff 'STOP'
   SymbolicIOField "Template_Symbolic I/O field_6" at 388,208 size 72x27; TextOn '1'; TextOff '0'; TextList "จัดเก็บ Motor speed1,2"
      ProcessValue <- "จัดเก็บ Servo DATA 1,2"
   SymbolicIOField "Template_Symbolic I/O field_7" at 388,238 size 72x27; TextOn '1'; TextOff '0'; TextList "จัดเก็บ Current 1,2"
      ProcessValue <- "จัดเก็บ Servo DATA 1,2"
   SymbolicIOField "Template_Symbolic I/O field_8" at 388,268 size 72x27; TextOn '1'; TextOff '0'; TextList "จัดเก็บ Power 1,2"
      ProcessValue <- "จัดเก็บ Servo DATA 1,2"
   SymbolicIOField "Template_Symbolic I/O field_9" at 388,298 size 72x27; TextOn '1'; TextOff '0'; TextList "จัดเก็บVoltage 1,2"
      ProcessValue <- "จัดเก็บ Servo DATA 1,2"
   SymbolicIOField "Template_Symbolic I/O field_10" at 637,208 size 72x27; TextOn '1'; TextOff '0'; TextList "จัดเก็บ Motor speed1,2"
      ProcessValue <- "จัดเก็บ Servo DATA 1,2"
   SymbolicIOField "Template_Symbolic I/O field_11" at 637,238 size 72x27; TextOn '1'; TextOff '0'; TextList "จัดเก็บ Current 1,2"
      ProcessValue <- "จัดเก็บ Servo DATA 1,2"
   SymbolicIOField "Template_Symbolic I/O field_12" at 636,269 size 72x27; TextOn '1'; TextOff '0'; TextList "จัดเก็บ Power 1,2"
      ProcessValue <- "จัดเก็บ Servo DATA 1,2"
   SymbolicIOField "Template_Symbolic I/O field_13" at 635,299 size 72x27; TextOn '1'; TextOff '0'; TextList "จัดเก็บVoltage 1,2"
      ProcessValue <- "จัดเก็บ Servo DATA 1,2"
   SymbolicIOField "Template_Symbolic I/O field_14" at 388,344 size 72x27; TextOn '1'; TextOff '0'; TextList "จัดเก็บ Motor speed3"
      ProcessValue <- "จัดเก็บ Servo DATA 3"
   SymbolicIOField "Template_Symbolic I/O field_15" at 388,373 size 72x27; TextOn '1'; TextOff '0'; TextList "จัดเก็บ Current 3"
      ProcessValue <- "จัดเก็บ Servo DATA 3"
   SymbolicIOField "Template_Symbolic I/O field_16" at 388,402 size 72x27; TextOn '1'; TextOff '0'; TextList "จัดเก็บ Power 3"
      ProcessValue <- "จัดเก็บ Servo DATA 3"
   SymbolicIOField "Template_Symbolic I/O field_17" at 388,431 size 72x27; TextOn '1'; TextOff '0'; TextList "จัดเก็บVoltage 3"
      ProcessValue <- "จัดเก็บ Servo DATA 3"
   GraphicView "Template_Graphic view_4" at 116,101 size 31x27; Picture "request"
   GraphicView "Template_Graphic view_5" at 176,293 size 24x24; Picture "add"
   GraphicView "Template_Graphic view_6" at 70,294 size 24x24; Picture "minus"
   GraphicView "Template_Graphic view_7" at 176,428 size 24x24; Picture "add"
   GraphicView "Template_Graphic view_8" at 70,429 size 24x24; Picture "minus"
   TextField "Template_Text field_10" at 294,213 size 99x17; Text 'Motor Speed 1'
   TextField "Template_Text field_11" at 459,213 size 30x17; Text 'rpm'
   TextField "Template_Text field_18" at 331,241 size 54x17; Text 'Current'
   TextField "Template_Text field_19" at 460,242 size 13x17; Text 'A'
   TextField "Template_Text field_21" at 338,271 size 44x17; Text 'Power'
   TextField "Template_Text field_22" at 459,272 size 16x17; Text 'W'
   TextField "Template_Text field_23" at 331,304 size 54x17; Text 'Voltage'
   TextField "Template_Text field_24" at 464,307 size 12x17; Text 'V'
   GraphicView "Template_Graphic view_1" at 185,100 size 39x35; Picture "box"
   GraphicView "Template_Graphic view_2" at 261,104 size 31x27; Picture "machine"
   GraphicView "Template_Graphic view_3" at 332,100 size 31x27; Picture "factory"
   TextField "Template_Text field_2" at 105,141 size 49x14; Text 'REQUEST'
   TextField "Template_Text field_12" at 192,142 size 28x14; Text 'PICK'
   TextField "Template_Text field_17" at 262,143 size 31x14; Text 'MOVE'
   TextField "Template_Text field_20" at 332,141 size 34x14; Text 'PLACE'
   TextField "Template_Text field_13" at 544,213 size 99x17; Text 'Motor Speed 2'
   TextField "Template_Text field_14" at 709,213 size 30x17; Text 'rpm'
   TextField "Template_Text field_15" at 581,241 size 54x17; Text 'Current'
   TextField "Template_Text field_16" at 710,242 size 13x17; Text 'A'
   TextField "Template_Text field_25" at 588,271 size 44x17; Text 'Power'
   TextField "Template_Text field_26" at 709,272 size 16x17; Text 'W'
   TextField "Template_Text field_27" at 581,304 size 54x17; Text 'Voltage'
   TextField "Template_Text field_28" at 714,307 size 12x17; Text 'V'
   TextField "Template_Text field_29" at 296,348 size 99x17; Text 'Motor Speed 3'
   TextField "Template_Text field_30" at 461,348 size 30x17; Text 'rpm'
   TextField "Template_Text field_31" at 333,376 size 54x17; Text 'Current'
   TextField "Template_Text field_32" at 462,377 size 13x17; Text 'A'
   TextField "Template_Text field_33" at 340,406 size 44x17; Text 'Power'
   TextField "Template_Text field_34" at 461,407 size 16x17; Text 'W'
   TextField "Template_Text field_35" at 333,439 size 54x17; Text 'Voltage'
   TextField "Template_Text field_36" at 466,442 size 12x17; Text 'V'
   TextField "Template_Text field_1" at 21,303 size 51x15; Text 'Encoder'
   TextField "Template_Text field_3" at 20,428 size 51x15; Text 'Encoder'
   TextField "Template_Text field_4" at 202,299 size 62x15; Text 'Pulse/rev'
   TextField "Template_Text field_5" at 201,432 size 62x15; Text 'Pulse/rev'
   TextField "Template_Text field_6" at 592,110 size 78x25; Text 'Storage'
   GraphicView "Template_Graphic view_9" at 437,92 size 54x52; Picture "KMUTNB-Photoroom"
   GraphicView "Template_Graphic view_10" at 470,82 size 126x131; Picture "MTET-Photoroom"
   Button "Button_1" at 177,294 size 24x24; TextOff 'Text'
   Button "Button_3" at 177,429 size 24x24; TextOff 'Text'
   Button "Button_2" at 70,295 size 24x24; TextOff 'Text'
   Button "Button_4" at 70,430 size 24x24; TextOff 'Text'

screen " propertyเบิกจ่าย" 800x480, template "property HMI data"
   SymbolicIOField "Template_Symbolic I/O field_2" at 19,248 size 122x32; TextOn '1'; TextOff '0'; TextList "X AXIS ( Horizontall )เบิกจ่าย"
      ProcessValue <- "แสดงชื่อยา"
   SymbolicIOField "Template_Symbolic I/O field_3" at 18,380 size 122x32; TextOn '1'; TextOff '0'; TextList "Y AXIS ( Verticall )เบิกจ่่าย"
      ProcessValue <- "แสดงชื่อยา"
   Circle "Template_Circle_5" at 104,87 size 56x56
      Appearance <- "รับคำสั่งเบิกยา"
   Circle "Template_Circle_2" at 252,88 size 56x56
      Appearance <- "Gripper หยิบยา"
   Circle "Template_Circle_4" at 180,87 size 56x56
      Appearance <- "เคลื่อนที่ไปยังตำยา"
   Circle "Template_Circle_7" at 320,87 size 56x56
      Appearance <- "เคลื่อนที่ไปยังตำแหน่งเริ่มต้น เบิกจ่าย"
   Button "Template_Button_2" at 688,88 size 96x64; TextOff 'Medicine Storage'
      on Press: ActivateScreen(" propertyจัดเก็บ", 0)
   Button "Template_Button_3" at 560,368 size 112x24; TextOff 'Reset to Default'
   Button "Template_Button_4" at 560,408 size 112x24; TextOff 'MODIFY'
   SymbolicIOField "Template_Symbolic I/O field_23" at 97,294 size 74x24; TextOn '1'; TextOff '0'; TextList "EncoderแกนX (เบิกจ่าย)"
      ProcessValue <- "แสดงชื่อยา"
   SymbolicIOField "Template_Symbolic I/O field_24" at 97,427 size 74x24; TextOn '1'; TextOff '0'; TextList "EncoderแกนY (เบิกจ่าย)"
      ProcessValue <- "แสดงชื่อยา"
   Button "Template_Button_1" at 681,422 size 88x24; TextOff 'HOME'
      on Press: ActivateScreen("1_OVERVIEW_1", 0)
   Button "Template_Button_5" at 681,358 size 88x24; TextOff 'START'
   Button "Template_Button_6" at 681,388 size 88x24; TextOff 'STOP'
   SymbolicIOField "Template_Symbolic I/O field_6" at 387,208 size 72x27; TextOn '1'; TextOff '0'; TextList "เบิกจ่าย Motor speed1,2"
      ProcessValue <- "เบิกจ่าย Servo DATA 1,2"
   SymbolicIOField "Template_Symbolic I/O field_7" at 387,238 size 72x27; TextOn '1'; TextOff '0'; TextList "เบิกจ่าย Current 1,2"
      ProcessValue <- "เบิกจ่าย Servo DATA 1,2"
   SymbolicIOField "Template_Symbolic I/O field_8" at 387,268 size 72x27; TextOn '1'; TextOff '0'; TextList "เบิกจ่าย Power 1,2"
      ProcessValue <- "เบิกจ่าย Servo DATA 1,2"
   SymbolicIOField "Template_Symbolic I/O field_9" at 387,298 size 72x27; TextOn '1'; TextOff '0'; TextList "เบิกจ่ายVoltage 1,2"
      ProcessValue <- "เบิกจ่าย Servo DATA 1,2"
   SymbolicIOField "Template_Symbolic I/O field_10" at 636,208 size 72x27; TextOn '1'; TextOff '0'; TextList "เบิกจ่าย Motor speed1,2"
      ProcessValue <- "เบิกจ่าย Servo DATA 1,2"
   SymbolicIOField "Template_Symbolic I/O field_11" at 636,238 size 72x27; TextOn '1'; TextOff '0'; TextList "เบิกจ่าย Current 1,2"
      ProcessValue <- "เบิกจ่าย Servo DATA 1,2"
   SymbolicIOField "Template_Symbolic I/O field_12" at 635,269 size 72x27; TextOn '1'; TextOff '0'; TextList "เบิกจ่าย Power 1,2"
      ProcessValue <- "เบิกจ่าย Servo DATA 1,2"
   SymbolicIOField "Template_Symbolic I/O field_13" at 634,299 size 72x27; TextOn '1'; TextOff '0'; TextList "เบิกจ่ายVoltage 1,2"
      ProcessValue <- "เบิกจ่าย Servo DATA 1,2"
   SymbolicIOField "Template_Symbolic I/O field_14" at 387,344 size 72x27; TextOn '1'; TextOff '0'; TextList "เบิกจ่าย Motor speed3"
      ProcessValue <- "เบิกจ่าย Servo DATA 3"
   SymbolicIOField "Template_Symbolic I/O field_15" at 387,373 size 72x27; TextOn '1'; TextOff '0'; TextList "เบิกจ่าย Current 3"
      ProcessValue <- "เบิกจ่าย Servo DATA 3"
   SymbolicIOField "Template_Symbolic I/O field_16" at 387,402 size 72x27; TextOn '1'; TextOff '0'; TextList "เบิกจ่าย Power 3"
      ProcessValue <- "เบิกจ่าย Servo DATA 3"
   SymbolicIOField "Template_Symbolic I/O field_17" at 387,431 size 72x27; TextOn '1'; TextOff '0'; TextList "เบิกจ่ายVoltage 3"
      ProcessValue <- "เบิกจ่าย Servo DATA 3"
   GraphicView "Template_Graphic view_4" at 116,101 size 31x27; Picture "request"
   GraphicView "Template_Graphic view_5" at 176,293 size 24x24; Picture "add"
   GraphicView "Template_Graphic view_6" at 70,294 size 24x24; Picture "minus"
   GraphicView "Template_Graphic view_7" at 175,426 size 24x24; Picture "add"
   GraphicView "Template_Graphic view_8" at 69,427 size 24x24; Picture "minus"
   TextField "Template_Text field_10" at 294,213 size 99x17; Text 'Motor Speed 1'
   TextField "Template_Text field_11" at 459,213 size 30x17; Text 'rpm'
   TextField "Template_Text field_18" at 331,241 size 54x17; Text 'Current'
   TextField "Template_Text field_19" at 460,242 size 13x17; Text 'A'
   TextField "Template_Text field_21" at 338,271 size 44x17; Text 'Power'
   TextField "Template_Text field_22" at 459,272 size 16x17; Text 'W'
   TextField "Template_Text field_23" at 331,304 size 54x17; Text 'Voltage'
   TextField "Template_Text field_24" at 464,307 size 12x17; Text 'V'
   GraphicView "Template_Graphic view_1" at 260,100 size 39x35; Picture "box"
   GraphicView "Template_Graphic view_2" at 193,103 size 31x27; Picture "machine"
   GraphicView "Template_Graphic view_3" at 332,100 size 31x27; Picture "factory"
   TextField "Template_Text field_2" at 105,141 size 49x14; Text 'REQUEST'
   TextField "Template_Text field_12" at 267,142 size 28x14; Text 'PICK'
   TextField "Template_Text field_17" at 194,142 size 31x14; Text 'MOVE'
   TextField "Template_Text field_20" at 332,141 size 34x14; Text 'PLACE'
   TextField "Template_Text field_13" at 544,213 size 99x17; Text 'Motor Speed 2'
   TextField "Template_Text field_14" at 709,213 size 30x17; Text 'rpm'
   TextField "Template_Text field_15" at 581,241 size 54x17; Text 'Current'
   TextField "Template_Text field_16" at 710,242 size 13x17; Text 'A'
   TextField "Template_Text field_25" at 588,271 size 44x17; Text 'Power'
   TextField "Template_Text field_26" at 709,272 size 16x17; Text 'W'
   TextField "Template_Text field_27" at 581,304 size 54x17; Text 'Voltage'
   TextField "Template_Text field_28" at 714,307 size 12x17; Text 'V'
   TextField "Template_Text field_29" at 296,348 size 99x17; Text 'Motor Speed 3'
   TextField "Template_Text field_30" at 461,348 size 30x17; Text 'rpm'
   TextField "Template_Text field_31" at 333,376 size 54x17; Text 'Current'
   TextField "Template_Text field_32" at 462,377 size 13x17; Text 'A'
   TextField "Template_Text field_33" at 340,406 size 44x17; Text 'Power'
   TextField "Template_Text field_34" at 461,407 size 16x17; Text 'W'
   TextField "Template_Text field_35" at 333,439 size 54x17; Text 'Voltage'
   TextField "Template_Text field_36" at 466,442 size 12x17; Text 'V'
   TextField "Template_Text field_1" at 21,298 size 51x15; Text 'Encoder'
   TextField "Template_Text field_3" at 20,431 size 51x15; Text 'Encoder'
   TextField "Template_Text field_4" at 202,298 size 61x15; Text 'Pulse/rev'
   TextField "Template_Text field_5" at 202,431 size 62x15; Text 'Pulse/rev'
   TextField "Template_Text field_6" at 594,106 size 89x25; Text 'Retrieval'
   GraphicView "Template_Graphic view_9" at 440,92 size 54x52; Picture "KMUTNB-Photoroom"
   GraphicView "Template_Graphic view_10" at 473,82 size 126x131; Picture "MTET-Photoroom"
   Button "Button_2" at 70,295 size 24x24; TextOff 'Text'
   Button "Button_3" at 69,428 size 24x24; TextOff 'Text'
   Button "Button_1" at 177,294 size 24x24; TextOff 'Text'
   Button "Button_4" at 176,427 size 24x24; TextOff 'Text'

screen "Status System" 800x480, template "Status system"
   Button "Button_3" at 666,441 size 120x36; TextOff 'Text'
      on Press: ActivateScreen("1_OVERVIEW_1", 0)
   Button "Button_1" at 545,441 size 120x36; TextOff 'Text'
      on Press: ActivateScreen("2_ALAREMS", 0)
   GraphicView "Template_Graphic view_5" at 678,446 size 24x25; Picture "NEW_HOME"
   TextField "Template_Text field_21" at 264,156 size 138x22; Text 'รับคำสั่งจัดเก็บยา'
   TextField "Template_Text field_24" at 275,244 size 118x40; Text 'เคลื่อนที่ไปยัง ตำแหน่งจัดเก็บ'
   TextField "Template_Text field_25" at 274,290 size 121x40; Text 'Gripper วางยา เข้าช่องจัดเก็บ'
   TextField "Template_Text field_26" at 277,337 size 118x40; Text 'เคลื่อนที่ไปยัง ตำแหน่งเริ่มต้น'
   TextField "Template_Text field_16" at 66,152 size 116x22; Text 'รับคำสั่งเบิกยา'
   TextField "Template_Text field_17" at 71,208 size 114x46; Text 'เคลื่อนที่ไปยังตำ แหน่งยา'
   TextField "Template_Text field_18" at 66,264 size 128x22; Text 'Gripper หยิบยา'
   TextField "Template_Text field_19" at 66,309 size 132x40; Text 'เคลื่อนที่ไปยังตำ แหน่งเริ่มต้น'
   TextField "Template_Text field_20" at 66,365 size 142x46; Text 'ยาไปช่องเบิกจ่าย / รอคำสั่งเบิกยา'
   TextField "Template_Text field_1" at 275,199 size 114x46; Text 'Gripperเคลื่อนที่ มารับยา'
   TextField "Template_Text field_2" at 280,390 size 142x22; Text 'รอรับคำสั่งยา'
   TextField "Text field_1" at 712,451 size 49x18; Text 'HOME'
   TextField "Text field_2" at 592,452 size 30x18; Text 'Doc'
   SymbolicIOField "Template_Symbolic I/O field_1" at 323,450 size 82x23; TextOn '1'; TextOff '0'
   SymbolicIOField "Template_Symbolic I/O field_2" at 120,450 size 82x23; TextOn '1'; TextOff '0'
   GraphicIOField "PlotLight_Square_G" at 230,146 size 42x42; PictureOff "PilotLight_Square_G_Off_256c"; PictureOn "PilotLight_Square_G_On_256c"
      ProcessValue <- "ป้อนรหัส Barcode"
   GraphicIOField "PlotLight_Square_G_1" at 230,195 size 42x42; PictureOn "PilotLight_Square_G_On_256c"; PictureOff "PilotLight_Square_G_Off_256c"
      ProcessValue <- "Gripperเคลื่อนที่มาเอายา"
   GraphicIOField "PlotLight_Square_G_2" at 230,242 size 42x42; PictureOn "PilotLight_Square_G_On_256c"; PictureOff "PilotLight_Square_G_Off_256c"
      ProcessValue <- "Gripper เคลื่อนไปช่องยา"
   GraphicIOField "PlotLight_Square_G_3" at 230,289 size 42x42; PictureOn "PilotLight_Square_G_On_256c"; PictureOff "PilotLight_Square_G_Off_256c"
      ProcessValue <- "Gripper วางยา"
   GraphicIOField "PlotLight_Square_G_4" at 230,336 size 42x42; PictureOn "PilotLight_Square_G_On_256c"; PictureOff "PilotLight_Square_G_Off_256c"
      ProcessValue <- "เคลื่อนที่ไปยังจุดเริ่มต้น"
   GraphicIOField "PlotLight_Square_G_5" at 230,383 size 42x42; PictureOn "PilotLight_Square_G_On_256c"; PictureOff "PilotLight_Square_G_Off_256c"
      ProcessValue <- "รอรับคำสั่งยา"
   GraphicIOField "PlotLight_Square_R" at 24,143 size 42x42; PictureOff "PilotLight_Square_R_Off_256c"; PictureOn "PilotLight_Square_R_On_256c"
      ProcessValue <- "รับคำสั่งเบิกยา"
   GraphicIOField "PlotLight_Square_R_1" at 23,201 size 42x42; PictureOn "PilotLight_Square_R_On_256c"; PictureOff "PilotLight_Square_R_Off_256c"
      ProcessValue <- "เคลื่อนที่ไปยังตำยา"
   GraphicIOField "PlotLight_Square_R_3" at 23,308 size 42x42; PictureOn "PilotLight_Square_R_On_256c"; PictureOff "PilotLight_Square_R_Off_256c"
      ProcessValue <- "เคลื่อนที่ไปยังตำแหน่งเริ่มต้น เบิกจ่าย"
   GraphicIOField "PlotLight_Square_R_4" at 23,363 size 42x42; PictureOn "PilotLight_Square_R_On_256c"; PictureOff "PilotLight_Square_R_Off_256c"
      ProcessValue <- "รอคำสั่งเบิกยา"
   TextField "Template_Text field_6" at 38,152 size 12x22; Text '1'
   TextField "Template_Text field_7" at 38,208 size 12x22; Text '2'
   TextField "Template_Text field_9" at 37,317 size 12x22; Text '4'
   TextField "Template_Text field_10" at 38,373 size 12x22; Text '5'
   TextField "Template_Text field_11" at 245,156 size 12x22; Text '1'
   TextField "Template_Text field_12" at 245,203 size 12x22; Text '2'
   TextField "Template_Text field_13" at 246,252 size 12x22; Text '3'
   TextField "Template_Text field_14" at 246,298 size 12x22; Text '4'
   TextField "Template_Text field_15" at 246,344 size 12x22; Text '5'
   TextField "Template_Text field_22" at 247,392 size 12x22; Text '6'
   GraphicIOField "PlotLight_Square_R_2" at 24,256 size 42x42; PictureOff "PilotLight_Square_R_Off_256c"; PictureOn "PilotLight_Square_R_On_256c"
      ProcessValue <- "Gripper หยิบยา"
   TextField "Template_Text field_3" at 40,264 size 12x22; Text '3'
   SymbolicIOField "Template_Symbolic I/O field_3" at 323,450 size 82x23; TextOn '1'; TextOff '0'; TextList "Status1"
      ProcessValue <- "Output Status1"
   SymbolicIOField "Template_Symbolic I/O field_4" at 120,450 size 82x23; TextOn '1'; TextOff '0'; TextList "Status1"
      ProcessValue <- "Output Status2"

screen "Screen_2" 800x480, template "Keep_1"
   Circle "Circle_2" at 38,164 size 32x32
      Appearance <- "Barcode46"
   Circle "Circle_1" at 38,224 size 32x32
      Appearance <- "Barcode55"
   Circle "Circle_3" at 38,279 size 32x32
      Appearance <- "Barcode64"
   Circle "Circle_4" at 38,336 size 32x32
      Appearance <- "Barcode73"
   Circle "Circle_5" at 38,393 size 32x32
      Appearance <- "Barcode82"
   Circle "Circle_6" at 102,164 size 32x32
      Appearance <- "Barcode47"
   Circle "Circle_7" at 102,224 size 32x32
      Appearance <- "Barcode56"
   Circle "Circle_8" at 102,279 size 32x32
      Appearance <- "Barcode65"
   Circle "Circle_9" at 102,336 size 32x32
      Appearance <- "Barcode74"
   Circle "Circle_10" at 102,393 size 32x32
      Appearance <- "Barcode83"
   Circle "Circle_11" at 166,164 size 32x32
      Appearance <- "Barcode48"
   Circle "Circle_12" at 166,224 size 32x32
      Appearance <- "Barcode57"
   Circle "Circle_13" at 166,279 size 32x32
      Appearance <- "Barcode66"
   Circle "Circle_14" at 166,336 size 32x32
      Appearance <- "Barcode75"
   Circle "Circle_15" at 166,393 size 32x32
      Appearance <- "Barcode84"
   Circle "Circle_16" at 230,164 size 32x32
      Appearance <- "Barcode49"
   Circle "Circle_17" at 230,224 size 32x32
      Appearance <- "Barcode58"
   Circle "Circle_18" at 230,279 size 32x32
      Appearance <- "Barcode67"
   Circle "Circle_19" at 230,336 size 32x32
      Appearance <- "Barcode76"
   Circle "Circle_20" at 230,393 size 32x32
      Appearance <- "Barcode85"
   Circle "Circle_21" at 294,164 size 32x32
      Appearance <- "Barcode50"
   Circle "Circle_22" at 294,224 size 32x32
      Appearance <- "Barcode59"
   Circle "Circle_23" at 294,279 size 32x32
      Appearance <- "Barcode68"
   Circle "Circle_24" at 294,336 size 32x32
      Appearance <- "Barcode77"
   Circle "Circle_25" at 294,393 size 32x32
      Appearance <- "Barcode86"
   Circle "Circle_26" at 358,164 size 32x32
      Appearance <- "Barcode51"
   Circle "Circle_27" at 358,225 size 32x32
      Appearance <- "Barcode60"
   Circle "Circle_28" at 358,279 size 32x32
      Appearance <- "Barcode69"
   Circle "Circle_29" at 358,336 size 32x32
      Appearance <- "Barcode78"
   Circle "Circle_30" at 358,393 size 32x32
      Appearance <- "Barcode87"
   Circle "Circle_31" at 422,164 size 32x32
      Appearance <- "Barcode52"
   Circle "Circle_32" at 422,224 size 32x32
      Appearance <- "Barcode61"
   Circle "Circle_33" at 422,279 size 32x32
      Appearance <- "Barcode70"
   Circle "Circle_34" at 422,336 size 32x32
      Appearance <- "Barcode79"
   Circle "Circle_35" at 422,393 size 32x32
      Appearance <- "Barcode88"
   Circle "Circle_36" at 486,164 size 32x32
      Appearance <- "Barcode53"
   Circle "Circle_37" at 486,224 size 32x32
      Appearance <- "Barcode62"
   Circle "Circle_38" at 486,279 size 32x32
      Appearance <- "Barcode71"
   Circle "Circle_39" at 486,336 size 32x32
      Appearance <- "Barcode80"
   Circle "Circle_40" at 486,393 size 32x32
      Appearance <- "Barcode89"
   Circle "Circle_41" at 550,163 size 32x32
      Appearance <- "Barcode54"
   Circle "Circle_42" at 550,224 size 32x32
      Appearance <- "Barcode63"
   Circle "Circle_43" at 550,279 size 32x32
      Appearance <- "Barcode72"
   Circle "Circle_44" at 550,336 size 32x32
      Appearance <- "Barcode81"
   Circle "Circle_45" at 550,393 size 32x32
      Appearance <- "Barcode90"
   TextField "Text field_1" at 30,146 size 57x20; Text 'Box_46'
   TextField "Text field_2" at 94,146 size 57x20; Text 'Box_47'
   TextField "Text field_3" at 159,146 size 57x20; Text 'Box_48'
   TextField "Text field_4" at 222,146 size 57x20; Text 'Box_49'
   TextField "Text field_5" at 286,146 size 57x20; Text 'Box_50'
   TextField "Text field_6" at 351,146 size 57x20; Text 'Box_51'
   TextField "Text field_7" at 415,146 size 57x20; Text 'Box_52'
   TextField "Text field_8" at 479,146 size 57x20; Text 'Box_53'
   TextField "Text field_9" at 542,146 size 57x20; Text 'Box_54'
   TextField "Text field_10" at 30,206 size 57x20; Text 'Box_55'
   TextField "Text field_11" at 92,206 size 57x20; Text 'Box_56'
   TextField "Text field_12" at 157,206 size 57x20; Text 'Box_57'
   TextField "Text field_13" at 222,206 size 57x20; Text 'Box_58'
   TextField "Text field_14" at 287,206 size 57x20; Text 'Box_59'
   TextField "Text field_15" at 350,206 size 57x20; Text 'Box_60'
   TextField "Text field_16" at 414,206 size 57x20; Text 'Box_61'
   TextField "Text field_17" at 478,206 size 57x20; Text 'Box_62'
   TextField "Text field_18" at 541,206 size 57x20; Text 'Box_63'
   TextField "Text field_19" at 31,261 size 57x20; Text 'Box_64'
   TextField "Text field_20" at 92,261 size 57x20; Text 'Box_65'
   TextField "Text field_21" at 157,261 size 57x20; Text 'Box_66'
   TextField "Text field_22" at 222,261 size 57x20; Text 'Box_67'
   TextField "Text field_23" at 287,261 size 57x20; Text 'Box_68'
   TextField "Text field_24" at 350,261 size 57x20; Text 'Box_69'
   TextField "Text field_25" at 414,261 size 57x20; Text 'Box_70'
   TextField "Text field_26" at 478,261 size 57x20; Text 'Box_71'
   TextField "Text field_27" at 541,261 size 57x20; Text 'Box_72'
   TextField "Text field_28" at 31,317 size 57x20; Text 'Box_73'
   TextField "Text field_29" at 92,317 size 57x20; Text 'Box_74'
   TextField "Text field_30" at 157,317 size 57x20; Text 'Box_75'
   TextField "Text field_31" at 222,317 size 57x20; Text 'Box_76'
   TextField "Text field_32" at 287,317 size 57x20; Text 'Box_77'
   TextField "Text field_33" at 350,317 size 57x20; Text 'Box_78'
   TextField "Text field_34" at 414,317 size 57x20; Text 'Box_79'
   TextField "Text field_35" at 478,317 size 57x20; Text 'Box_80'
   TextField "Text field_36" at 541,317 size 57x20; Text 'Box_81'
   TextField "Text field_37" at 31,375 size 57x20; Text 'Box_82'
   TextField "Text field_38" at 92,375 size 57x20; Text 'Box_83'
   TextField "Text field_39" at 157,375 size 57x20; Text 'Box_84'
   TextField "Text field_40" at 222,375 size 57x20; Text 'Box_85'
   TextField "Text field_41" at 287,375 size 57x20; Text 'Box_86'
   TextField "Text field_42" at 350,375 size 57x20; Text 'Box_87'
   TextField "Text field_43" at 414,375 size 57x20; Text 'Box_88'
   TextField "Text field_44" at 478,375 size 57x20; Text 'Box_89'
   TextField "Text field_45" at 541,375 size 57x20; Text 'Box_90'
   SymbolicIOField "Symbolic I/O field_1" at 621,342 size 167x24; TextOn '1'; TextOff '0'; TextList "BOX_All"
      ProcessValue <- "แสดงชื่อยา2"
   IOField "I/O field_1" at 624,160 size 160x64; FormatPattern ???????????
      on OnFinishInput: "Test2"(); "Storage"()
      ProcessValue <- "Expected/Value_All_V"
   TextField "Text field_47" at 648,418 size 78x17; Text ': Low Stock'
   TextField "Text field_46" at 646,395 size 104x17; Text ': Medium Stock'
   TextField "Text field_48" at 646,372 size 82x17; Text ': High Stock'
   Button "Button_5" at 633,292 size 64x24; TextOff 'Back'
      on Click: ActivateScreen("Screen_1", 0)
   Button "Button_6" at 716,292 size 64x24; TextOff 'Next'
      on Click: ActivateScreen("Screen_3", 0)
   GraphicView "Template_Graphic view_1" at 16,8 size 70x68; Picture "KMUTNB-Photoroom"
   GraphicView "Template_Graphic view_5" at 657,59 size 104x124; Picture "channels4_profile-Photoroom"
   GraphicView "Template_Graphic view_2" at 736,255 size 28x26; Picture "NEW_HOME"
   GraphicView "Template_Graphic view_6" at 650,253 size 28x27; Picture "play"
   GraphicView "Template_Graphic view_3" at 721,296 size 20x17; Picture "next-track"
   GraphicView "Template_Graphic view_4" at 638,296 size 20x17; Picture "previous-track"
   Button "Button_3" at 707,246 size 80x42; TextOn 'LOGOUT'; TextOff 'Text'
      on Activate: function_f23ef4c9(); ActivateScreen("1_OVERVIEW_1", 0)
   Button "Button_1" at 623,245 size 80x42; TextOff 'Text'
      on Press: SetTag("มีการปุ่มกดยืนยัน", 1)
      on Release: SetTag("มีการปุ่มกดยืนยัน", 0)
      on Activate: "Storage"()
      on Click: "Conveyor"(); ActivateScreen("Status System", 0)
   TextField "Text field_49" at 734,229 size 32x14; Text 'HOME'
   TextField "Text field_50" at 625,229 size 95x16; Text 'Simmulation Conveyor'

screen "LOGIN_1" 800x480, template "Template"
   Button "Button_2" at 668,96 size 128x72; TextOff 'LOGIN'; Authorization "Admin"
      on Activate: function_a2a04561(); ActivateScreen("Screen_1", 0)
   Button "Button_6" at 668,398 size 128x72; TextOn 'LOGOUT'; TextOff 'LOGOUT'
      on Activate: function_f23ef4c9(); ActivateScreen("1_OVERVIEW_1", 0)
   GraphicView "Template_Graphic view_1" at 672,107 size 54x48; Picture "NEW_HOME"
   GraphicView "Template_Graphic view_5" at 672,413 size 54x48; Picture "logout"

screen "Screen_1" 800x480, template "Keep_1"
   IOField "I/O field_1" at 624,160 size 160x64; FormatPattern ???????????
      on OnFinishInput: "Storage"()
      ProcessValue <- "Expected/Value_All_V"
   TextField "Text field_1" at 35,146 size 48x20; Text 'Box_1'
   TextField "Text field_2" at 96,146 size 48x20; Text 'Box_2'
   TextField "Text field_3" at 161,146 size 48x20; Text 'Box_3'
   TextField "Text field_4" at 226,146 size 48x20; Text 'Box_4'
   TextField "Text field_5" at 291,146 size 48x20; Text 'Box_5'
   TextField "Text field_6" at 354,146 size 48x20; Text 'Box_6'
   TextField "Text field_7" at 418,146 size 48x20; Text 'Box_7'
   TextField "Text field_8" at 482,146 size 48x20; Text 'Box_8'
   TextField "Text field_9" at 545,146 size 48x20; Text 'Box_9'
   TextField "Text field_10" at 31,206 size 57x20; Text 'Box_10'
   TextField "Text field_11" at 92,206 size 57x20; Text 'Box_11'
   TextField "Text field_12" at 157,206 size 57x20; Text 'Box_12'
   TextField "Text field_13" at 222,206 size 57x20; Text 'Box_13'
   TextField "Text field_14" at 287,206 size 57x20; Text 'Box_14'
   TextField "Text field_15" at 350,206 size 57x20; Text 'Box_15'
   TextField "Text field_16" at 414,206 size 57x20; Text 'Box_16'
   TextField "Text field_17" at 478,206 size 57x20; Text 'Box_17'
   TextField "Text field_18" at 541,206 size 57x20; Text 'Box_18'
   TextField "Text field_19" at 31,261 size 57x20; Text 'Box_19'
   TextField "Text field_20" at 92,261 size 57x20; Text 'Box_20'
   TextField "Text field_21" at 157,261 size 57x20; Text 'Box_21'
   TextField "Text field_22" at 222,261 size 57x20; Text 'Box_22'
   TextField "Text field_23" at 287,261 size 57x20; Text 'Box_23'
   TextField "Text field_24" at 350,261 size 57x20; Text 'Box_24'
   TextField "Text field_25" at 414,261 size 57x20; Text 'Box_25'
   TextField "Text field_26" at 478,261 size 57x20; Text 'Box_26'
   TextField "Text field_27" at 541,261 size 57x20; Text 'Box_27'
   TextField "Text field_28" at 31,317 size 57x20; Text 'Box_28'
   TextField "Text field_29" at 92,317 size 57x20; Text 'Box_29'
   TextField "Text field_30" at 157,317 size 57x20; Text 'Box_30'
   TextField "Text field_31" at 222,317 size 57x20; Text 'Box_31'
   TextField "Text field_32" at 287,317 size 57x20; Text 'Box_32'
   TextField "Text field_33" at 350,317 size 57x20; Text 'Box_33'
   TextField "Text field_34" at 414,317 size 57x20; Text 'Box_34'
   TextField "Text field_35" at 478,317 size 57x20; Text 'Box_35'
   TextField "Text field_36" at 541,317 size 57x20; Text 'Box_36'
   TextField "Text field_37" at 31,375 size 57x20; Text 'Box_37'
   TextField "Text field_38" at 92,375 size 57x20; Text 'Box_38'
   TextField "Text field_39" at 157,375 size 57x20; Text 'Box_39'
   TextField "Text field_40" at 222,375 size 57x20; Text 'Box_40'
   TextField "Text field_41" at 287,375 size 57x20; Text 'Box_41'
   TextField "Text field_42" at 350,375 size 57x20; Text 'Box_42'
   TextField "Text field_43" at 414,375 size 57x20; Text 'Box_43'
   TextField "Text field_44" at 478,375 size 57x20; Text 'Box_44'
   TextField "Text field_45" at 541,375 size 57x20; Text 'Box_45'
   SymbolicIOField "Symbolic I/O field_1" at 621,342 size 167x24; TextOn '1'; TextOff '0'; TextList "BOX_All"
      ProcessValue <- "แสดงชื่อยา2"
   TextField "Text field_47" at 648,418 size 78x17; Text ': Low Stock'
   TextField "Text field_46" at 646,395 size 104x17; Text ': Medium Stock'
   TextField "Text field_48" at 646,372 size 82x17; Text ': High Stock'
   Circle "Circle_2" at 38,164 size 32x32
      Appearance <- "Barcode1"
   Circle "Circle_1" at 38,224 size 32x32
      Appearance <- "Barcode10"
   Circle "Circle_3" at 38,279 size 32x32
      Appearance <- "Barcode19"
   Circle "Circle_4" at 38,336 size 32x32
      Appearance <- "Barcode28"
   Circle "Circle_5" at 38,393 size 32x32
      Appearance <- "Barcode37"
   Circle "Circle_6" at 102,164 size 32x32
      Appearance <- "Barcode2"
   Circle "Circle_7" at 102,224 size 32x32
      Appearance <- "Barcode11"
   Circle "Circle_8" at 102,279 size 32x32
      Appearance <- "Barcode20"
   Circle "Circle_9" at 102,336 size 32x32
      Appearance <- "Barcode29"
   Circle "Circle_10" at 102,393 size 32x32
      Appearance <- "Barcode38"
   Circle "Circle_11" at 166,164 size 32x32
      Appearance <- "Barcode3"
   Circle "Circle_12" at 166,224 size 32x32
      Appearance <- "Barcode12"
   Circle "Circle_13" at 166,279 size 32x32
      Appearance <- "Barcode21"
   Circle "Circle_14" at 166,336 size 32x32
      Appearance <- "Barcode30"
   Circle "Circle_15" at 166,393 size 32x32
      Appearance <- "Barcode39"
   Circle "Circle_16" at 230,164 size 32x32
      Appearance <- "Barcode4"
   Circle "Circle_17" at 230,224 size 32x32
      Appearance <- "Barcode13"
   Circle "Circle_18" at 230,279 size 32x32
      Appearance <- "Barcode22"
   Circle "Circle_19" at 230,336 size 32x32
      Appearance <- "Barcode31"
   Circle "Circle_20" at 230,393 size 32x32
      Appearance <- "Barcode40"
   Circle "Circle_21" at 294,164 size 32x32
      Appearance <- "Barcode5"
   Circle "Circle_22" at 294,224 size 32x32
      Appearance <- "Barcode14"
   Circle "Circle_23" at 294,279 size 32x32
      Appearance <- "Barcode23"
   Circle "Circle_24" at 294,336 size 32x32
      Appearance <- "Barcode32"
   Circle "Circle_25" at 294,393 size 32x32
      Appearance <- "Barcode41"
   Circle "Circle_26" at 358,164 size 32x32
      Appearance <- "Barcode6"
   Circle "Circle_27" at 358,225 size 32x32
      Appearance <- "Barcode15"
   Circle "Circle_28" at 358,279 size 32x32
      Appearance <- "Barcode24"
   Circle "Circle_29" at 358,336 size 32x32
      Appearance <- "Barcode33"
   Circle "Circle_30" at 358,393 size 32x32
      Appearance <- "Barcode42"
   Circle "Circle_31" at 422,164 size 32x32
      Appearance <- "Barcode7"
   Circle "Circle_32" at 422,224 size 32x32
      Appearance <- "Barcode16"
   Circle "Circle_33" at 422,279 size 32x32
      Appearance <- "Barcode25"
   Circle "Circle_34" at 422,336 size 32x32
      Appearance <- "Barcode34"
   Circle "Circle_35" at 422,393 size 32x32
      Appearance <- "Barcode43"
   Circle "Circle_36" at 486,164 size 32x32
      Appearance <- "Barcode8"
   Circle "Circle_37" at 486,224 size 32x32
      Appearance <- "Barcode17"
   Circle "Circle_38" at 486,279 size 32x32
      Appearance <- "Barcode26"
   Circle "Circle_39" at 486,336 size 32x32
      Appearance <- "Barcode35"
   Circle "Circle_40" at 486,393 size 32x32
      Appearance <- "Barcode44"
   Circle "Circle_41" at 550,163 size 32x32
      Appearance <- "Barcode9"
   Circle "Circle_42" at 550,224 size 32x32
      Appearance <- "Barcode18"
   Circle "Circle_43" at 550,279 size 32x32
      Appearance <- "Barcode27"
   Circle "Circle_44" at 550,336 size 32x32
      Appearance <- "Barcode36"
   Circle "Circle_45" at 550,393 size 32x32
      Appearance <- "Barcode45"
   Button "Button_1" at 623,245 size 80x42; TextOff 'Text'
      on Click: "Conveyor"(); ActivateScreen("Status System", 0)
      on Activate: "Storage"()
      on Release: SetTag("มีการปุ่มกดยืนยัน", 0)
      on Press: SetTag("มีการปุ่มกดยืนยัน", 1)
   Button "Button_3" at 707,246 size 80x42; TextOn 'LOGOUT'; TextOff 'Text'
      on Activate: function_f23ef4c9(); ActivateScreen("1_OVERVIEW_1", 0)
   GraphicView "Template_Graphic view_3" at 721,296 size 20x17; Picture "next-track"
   GraphicView "Template_Graphic view_5" at 657,59 size 104x124; Picture "channels4_profile-Photoroom"
   Button "Button_6" at 716,292 size 64x24; TextOff 'Next'
      on Click: ActivateScreen("Screen_2", 0)
   GraphicView "Template_Graphic view_4" at 736,255 size 28x26; Picture "NEW_HOME"
   GraphicView "Template_Graphic view_1" at 16,8 size 70x68; Picture "KMUTNB-Photoroom"
   GraphicView "Template_Graphic view_2" at 650,253 size 28x27; Picture "play"
   TextField "Text field_49" at 734,229 size 32x14; Text 'HOME'
   TextField "Text field_50" at 625,229 size 95x16; Text 'Simmulation Conveyor'

screen "Screen_3" 800x480, template "Keep_1"
   TextField "Text field_1" at 32,146 size 57x20; Text 'Box_91'
   TextField "Text field_2" at 93,146 size 57x20; Text 'Box_92'
   TextField "Text field_3" at 158,146 size 57x20; Text 'Box_93'
   TextField "Text field_4" at 223,146 size 57x20; Text 'Box_94'
   TextField "Text field_5" at 288,146 size 57x20; Text 'Box_95'
   TextField "Text field_6" at 351,146 size 57x20; Text 'Box_96'
   TextField "Text field_7" at 415,146 size 57x20; Text 'Box_97'
   TextField "Text field_8" at 479,146 size 57x20; Text 'Box_98'
   TextField "Text field_9" at 542,146 size 57x20; Text 'Box_99'
   TextField "Text field_10" at 25,206 size 66x20; Text 'Box_100'
   TextField "Text field_11" at 88,206 size 66x20; Text 'Box_101'
   TextField "Text field_12" at 153,206 size 66x20; Text 'Box_102'
   TextField "Text field_13" at 217,206 size 66x20; Text 'Box_103'
   TextField "Text field_14" at 281,206 size 66x20; Text 'Box_104'
   TextField "Text field_15" at 345,206 size 66x20; Text 'Box_105'
   TextField "Text field_16" at 410,206 size 66x20; Text 'Box_106'
   TextField "Text field_17" at 473,206 size 66x20; Text 'Box_107'
   TextField "Text field_18" at 537,206 size 66x20; Text 'Box_108'
   TextField "Text field_19" at 26,261 size 66x20; Text 'Box_109'
   TextField "Text field_20" at 89,261 size 66x20; Text 'Box_110'
   TextField "Text field_21" at 153,261 size 66x20; Text 'Box_111'
   TextField "Text field_22" at 217,261 size 66x20; Text 'Box_112'
   TextField "Text field_23" at 281,261 size 66x20; Text 'Box_113'
   TextField "Text field_24" at 346,261 size 66x20; Text 'Box_114'
   TextField "Text field_25" at 409,261 size 66x20; Text 'Box_115'
   TextField "Text field_26" at 473,261 size 66x20; Text 'Box_116'
   TextField "Text field_27" at 537,261 size 66x20; Text 'Box_117'
   TextField "Text field_28" at 25,317 size 66x20; Text 'Box_118'
   TextField "Text field_29" at 88,317 size 66x20; Text 'Box_119'
   TextField "Text field_30" at 153,317 size 66x20; Text 'Box_120'
   TextField "Text field_31" at 218,317 size 66x20; Text 'Box_121'
   TextField "Text field_32" at 282,317 size 66x20; Text 'Box_122'
   TextField "Text field_33" at 346,317 size 66x20; Text 'Box_123'
   TextField "Text field_34" at 410,317 size 66x20; Text 'Box_124'
   TextField "Text field_35" at 472,317 size 66x20; Text 'Box_125'
   TextField "Text field_36" at 537,317 size 66x20; Text 'Box_126'
   TextField "Text field_37" at 26,375 size 66x20; Text 'Box_127'
   TextField "Text field_38" at 88,375 size 66x20; Text 'Box_128'
   TextField "Text field_39" at 153,375 size 66x20; Text 'Box_129'
   TextField "Text field_40" at 217,375 size 66x20; Text 'Box_130'
   TextField "Text field_41" at 281,375 size 66x20; Text 'Box_131'
   TextField "Text field_42" at 345,375 size 66x20; Text 'Box_132'
   TextField "Text field_43" at 409,375 size 66x20; Text 'Box_133'
   TextField "Text field_44" at 473,375 size 66x20; Text 'Box_134'
   TextField "Text field_45" at 536,375 size 66x20; Text 'Box_135'
   SymbolicIOField "Symbolic I/O field_1" at 621,342 size 167x24; TextOn '1'; TextOff '0'; TextList "BOX_All"
      ProcessValue <- "แสดงชื่อยา2"
   IOField "I/O field_1" at 624,160 size 160x64; FormatPattern ???????????
      on OnFinishInput: "Test2"(); "Storage"()
      ProcessValue <- "Expected/Value_All_V"
   TextField "Text field_47" at 648,418 size 78x17; Text ': Low Stock'
   TextField "Text field_46" at 646,395 size 104x17; Text ': Medium Stock'
   TextField "Text field_48" at 646,372 size 82x17; Text ': High Stock'
   Circle "Circle_2" at 38,164 size 32x32
      Appearance <- "Barcode91"
   Circle "Circle_1" at 38,224 size 32x32
      Appearance <- "Barcode100"
   Circle "Circle_3" at 38,279 size 32x32
      Appearance <- "Barcode109"
   Circle "Circle_4" at 38,336 size 32x32
      Appearance <- "Barcode118"
   Circle "Circle_5" at 38,393 size 32x32
      Appearance <- "Barcode127"
   Circle "Circle_6" at 102,164 size 32x32
      Appearance <- "Barcode92"
   Circle "Circle_7" at 102,224 size 32x32
      Appearance <- "Barcode101"
   Circle "Circle_8" at 102,279 size 32x32
      Appearance <- "Barcode110"
   Circle "Circle_9" at 102,336 size 32x32
      Appearance <- "Barcode119"
   Circle "Circle_10" at 102,393 size 32x32
      Appearance <- "Barcode128"
   Circle "Circle_11" at 166,164 size 32x32
      Appearance <- "Barcode93"
   Circle "Circle_12" at 166,224 size 32x32
      Appearance <- "Barcode102"
   Circle "Circle_13" at 166,279 size 32x32
      Appearance <- "Barcode111"
   Circle "Circle_14" at 166,336 size 32x32
      Appearance <- "Barcode120"
   Circle "Circle_15" at 166,393 size 32x32
      Appearance <- "Barcode129"
   Circle "Circle_16" at 230,164 size 32x32
      Appearance <- "Barcode94"
   Circle "Circle_17" at 230,224 size 32x32
      Appearance <- "Barcode103"
   Circle "Circle_18" at 230,279 size 32x32
      Appearance <- "Barcode112"
   Circle "Circle_19" at 230,336 size 32x32
      Appearance <- "Barcode121"
   Circle "Circle_20" at 230,393 size 32x32
      Appearance <- "Barcode130"
   Circle "Circle_21" at 294,164 size 32x32
      Appearance <- "Barcode95"
   Circle "Circle_22" at 294,224 size 32x32
      Appearance <- "Barcode104"
   Circle "Circle_23" at 294,279 size 32x32
      Appearance <- "Barcode113"
   Circle "Circle_24" at 294,336 size 32x32
      Appearance <- "Barcode122"
   Circle "Circle_25" at 294,393 size 32x32
      Appearance <- "Barcode131"
   Circle "Circle_26" at 358,164 size 32x32
      Appearance <- "Barcode96"
   Circle "Circle_27" at 358,225 size 32x32
      Appearance <- "Barcode105"
   Circle "Circle_28" at 358,279 size 32x32
      Appearance <- "Barcode114"
   Circle "Circle_29" at 358,336 size 32x32
      Appearance <- "Barcode123"
   Circle "Circle_30" at 358,393 size 32x32
      Appearance <- "Barcode132"
   Circle "Circle_31" at 422,164 size 32x32
      Appearance <- "Barcode97"
   Circle "Circle_32" at 422,224 size 32x32
      Appearance <- "Barcode106"
   Circle "Circle_33" at 422,279 size 32x32
      Appearance <- "Barcode115"
   Circle "Circle_34" at 422,336 size 32x32
      Appearance <- "Barcode124"
   Circle "Circle_35" at 422,393 size 32x32
      Appearance <- "Barcode133"
   Circle "Circle_36" at 486,164 size 32x32
      Appearance <- "Barcode98"
   Circle "Circle_37" at 486,224 size 32x32
      Appearance <- "Barcode107"
   Circle "Circle_38" at 486,279 size 32x32
      Appearance <- "Barcode116"
   Circle "Circle_39" at 486,336 size 32x32
      Appearance <- "Barcode125"
   Circle "Circle_40" at 486,393 size 32x32
      Appearance <- "Barcode134"
   Circle "Circle_41" at 550,163 size 32x32
      Appearance <- "Barcode99"
   Circle "Circle_42" at 550,224 size 32x32
      Appearance <- "Barcode108"
   Circle "Circle_43" at 550,279 size 32x32
      Appearance <- "Barcode117"
   Circle "Circle_44" at 550,336 size 32x32
      Appearance <- "Barcode126"
   Circle "Circle_45" at 550,393 size 32x32
      Appearance <- "Barcode135"
   GraphicView "Template_Graphic view_6" at 16,8 size 70x68; Picture "KMUTNB-Photoroom"
   GraphicView "Template_Graphic view_5" at 657,59 size 104x124; Picture "channels4_profile-Photoroom"
   Button "Button_5" at 633,292 size 64x24; TextOff 'Back'
      on Click: ActivateScreen("Screen_2", 0)
   Button "Button_6" at 716,292 size 64x24; TextOff 'Next'
      on Click: ActivateScreen("Screen_4", 0)
   GraphicView "Template_Graphic view_1" at 736,255 size 28x26; Picture "NEW_HOME"
   GraphicView "Template_Graphic view_2" at 650,253 size 28x27; Picture "play"
   GraphicView "Template_Graphic view_3" at 721,296 size 20x17; Picture "next-track"
   GraphicView "Template_Graphic view_4" at 638,296 size 20x17; Picture "previous-track"
   Button "Button_3" at 707,246 size 80x42; TextOn 'LOGOUT'; TextOff 'Text'
      on Activate: function_f23ef4c9(); ActivateScreen("1_OVERVIEW_1", 0)
   Button "Button_1" at 623,245 size 80x42; TextOff 'Text'
      on Press: SetTag("มีการปุ่มกดยืนยัน", 1)
      on Release: SetTag("มีการปุ่มกดยืนยัน", 0)
      on Activate: "Storage"()
      on Click: "Conveyor"(); ActivateScreen("Status System", 0)
   TextField "Text field_49" at 734,229 size 32x14; Text 'HOME'
   TextField "Text field_50" at 625,229 size 95x16; Text 'Simmulation Conveyor'

screen "Screen_4" 800x480, template "Keep_1"
   Circle "Circle_2" at 38,164 size 32x32
      Appearance <- "Barcode136"
   Circle "Circle_1" at 38,224 size 32x32
      Appearance <- "Barcode145"
   Circle "Circle_3" at 38,279 size 32x32
      Appearance <- "Barcode154"
   Circle "Circle_4" at 38,336 size 32x32
      Appearance <- "Barcode163"
   Circle "Circle_5" at 38,393 size 32x32
      Appearance <- "Barcode172"
   Circle "Circle_6" at 102,164 size 32x32
      Appearance <- "Barcode137"
   Circle "Circle_7" at 102,224 size 32x32
      Appearance <- "Barcode146"
   Circle "Circle_8" at 102,279 size 32x32
      Appearance <- "Barcode155"
   Circle "Circle_9" at 102,336 size 32x32
      Appearance <- "Barcode164"
   Circle "Circle_10" at 102,393 size 32x32
      Appearance <- "Barcode173"
   Circle "Circle_11" at 166,164 size 32x32
      Appearance <- "Barcode138"
   Circle "Circle_12" at 166,224 size 32x32
      Appearance <- "Barcode147"
   Circle "Circle_13" at 166,279 size 32x32
      Appearance <- "Barcode156"
   Circle "Circle_14" at 166,336 size 32x32
      Appearance <- "Barcode165"
   Circle "Circle_15" at 166,393 size 32x32
      Appearance <- "Barcode174"
   Circle "Circle_16" at 230,164 size 32x32
      Appearance <- "Barcode139"
   Circle "Circle_17" at 230,224 size 32x32
      Appearance <- "Barcode148"
   Circle "Circle_18" at 230,279 size 32x32
      Appearance <- "Barcode157"
   Circle "Circle_19" at 230,336 size 32x32
      Appearance <- "Barcode166"
   Circle "Circle_20" at 230,393 size 32x32
      Appearance <- "Barcode175"
   Circle "Circle_21" at 294,164 size 32x32
      Appearance <- "Barcode140"
   Circle "Circle_22" at 294,224 size 32x32
      Appearance <- "Barcode149"
   Circle "Circle_23" at 294,279 size 32x32
      Appearance <- "Barcode158"
   Circle "Circle_24" at 294,336 size 32x32
      Appearance <- "Barcode167"
   Circle "Circle_25" at 294,393 size 32x32
      Appearance <- "Barcode176"
   Circle "Circle_26" at 358,164 size 32x32
      Appearance <- "Barcode141"
   Circle "Circle_27" at 358,225 size 32x32
      Appearance <- "Barcode150"
   Circle "Circle_28" at 358,279 size 32x32
      Appearance <- "Barcode159"
   Circle "Circle_29" at 358,336 size 32x32
      Appearance <- "Barcode168"
   Circle "Circle_30" at 358,393 size 32x32
      Appearance <- "Barcode177"
   Circle "Circle_31" at 422,164 size 32x32
      Appearance <- "Barcode142"
   Circle "Circle_32" at 422,224 size 32x32
      Appearance <- "Barcode151"
   Circle "Circle_33" at 422,279 size 32x32
      Appearance <- "Barcode160"
   Circle "Circle_34" at 422,336 size 32x32
      Appearance <- "Barcode169"
   Circle "Circle_35" at 422,393 size 32x32
      Appearance <- "Barcode178"
   Circle "Circle_36" at 486,164 size 32x32
      Appearance <- "Barcode143"
   Circle "Circle_37" at 486,224 size 32x32
      Appearance <- "Barcode152"
   Circle "Circle_38" at 486,279 size 32x32
      Appearance <- "Barcode161"
   Circle "Circle_39" at 486,336 size 32x32
      Appearance <- "Barcode170"
   Circle "Circle_40" at 486,393 size 32x32
      Appearance <- "Barcode179"
   Circle "Circle_41" at 550,163 size 32x32
      Appearance <- "Barcode144"
   Circle "Circle_42" at 550,224 size 32x32
      Appearance <- "Barcode153"
   Circle "Circle_43" at 550,279 size 32x32
      Appearance <- "Barcode162"
   Circle "Circle_44" at 550,336 size 32x32
      Appearance <- "Barcode171"
   Circle "Circle_45" at 550,393 size 32x32
      Appearance <- "Barcode180"
   TextField "Text field_8" at 473,145 size 66x20; Text 'Box_143'
   TextField "Text field_9" at 536,145 size 66x20; Text 'Box_144'
   TextField "Text field_10" at 25,206 size 66x20; Text 'Box_145'
   TextField "Text field_11" at 88,206 size 66x20; Text 'Box_146'
   TextField "Text field_12" at 153,206 size 66x20; Text 'Box_147'
   TextField "Text field_13" at 217,206 size 66x20; Text 'Box_148'
   TextField "Text field_14" at 281,206 size 66x20; Text 'Box_149'
   TextField "Text field_15" at 345,206 size 66x20; Text 'Box_150'
   TextField "Text field_16" at 410,206 size 66x20; Text 'Box_151'
   TextField "Text field_17" at 473,206 size 66x20; Text 'Box_152'
   TextField "Text field_19" at 26,261 size 66x20; Text 'Box_154'
   TextField "Text field_20" at 89,261 size 66x20; Text 'Box_155'
   TextField "Text field_21" at 153,261 size 66x20; Text 'Box_156'
   TextField "Text field_22" at 217,261 size 66x20; Text 'Box_157'
   TextField "Text field_23" at 281,261 size 66x20; Text 'Box_158'
   TextField "Text field_24" at 346,261 size 66x20; Text 'Box_159'
   TextField "Text field_25" at 409,261 size 66x20; Text 'Box_160'
   TextField "Text field_26" at 473,261 size 66x20; Text 'Box_161'
   TextField "Text field_28" at 25,317 size 66x20; Text 'Box_163'
   TextField "Text field_29" at 88,317 size 66x20; Text 'Box_164'
   TextField "Text field_30" at 153,317 size 66x20; Text 'Box_165'
   TextField "Text field_31" at 218,317 size 66x20; Text 'Box_166'
   TextField "Text field_32" at 282,317 size 66x20; Text 'Box_167'
   TextField "Text field_33" at 346,317 size 66x20; Text 'Box_168'
   TextField "Text field_34" at 410,317 size 66x20; Text 'Box_169'
   TextField "Text field_35" at 472,317 size 66x20; Text 'Box_170'
   TextField "Text field_37" at 26,375 size 66x20; Text 'Box_172'
   TextField "Text field_38" at 88,375 size 66x20; Text 'Box_173'
   TextField "Text field_39" at 153,375 size 66x20; Text 'Box_174'
   TextField "Text field_40" at 217,375 size 66x20; Text 'Box_175'
   TextField "Text field_41" at 281,375 size 66x20; Text 'Box_176'
   TextField "Text field_42" at 345,375 size 66x20; Text 'Box_177'
   TextField "Text field_43" at 409,375 size 66x20; Text 'Box_178'
   TextField "Text field_44" at 473,375 size 66x20; Text 'Box_179'
   TextField "Text field_18" at 537,206 size 66x20; Text 'Box_153'
   TextField "Text field_27" at 537,261 size 66x20; Text 'Box_162'
   TextField "Text field_36" at 537,317 size 66x20; Text 'Box_171'
   TextField "Text field_45" at 536,375 size 66x20; Text 'Box_180'
   TextField "Text field_1" at 24,145 size 66x20; Text 'Box_136'
   TextField "Text field_2" at 87,145 size 66x20; Text 'Box_137'
   TextField "Text field_3" at 152,145 size 66x20; Text 'Box_138'
   TextField "Text field_4" at 216,145 size 66x20; Text 'Box_139'
   TextField "Text field_5" at 280,145 size 66x20; Text 'Box_140'
   TextField "Text field_6" at 344,145 size 66x20; Text 'Box_141'
   TextField "Text field_7" at 409,145 size 66x20; Text 'Box_142'
   SymbolicIOField "Symbolic I/O field_1" at 621,342 size 167x24; TextOn '1'; TextOff '0'; TextList "BOX_All"
      ProcessValue <- "แสดงชื่อยา2"
   IOField "I/O field_1" at 624,160 size 160x64; FormatPattern ???????????
      on OnFinishInput: "Test2"(); "Storage"()
      ProcessValue <- "Expected/Value_All_V"
   TextField "Text field_47" at 648,418 size 78x17; Text ': Low Stock'
   TextField "Text field_46" at 646,395 size 104x17; Text ': Medium Stock'
   TextField "Text field_48" at 646,372 size 82x17; Text ': High Stock'
   GraphicView "Template_Graphic view_6" at 16,8 size 70x68; Picture "KMUTNB-Photoroom"
   GraphicView "Template_Graphic view_5" at 657,59 size 104x124; Picture "channels4_profile-Photoroom"
   Button "Button_5" at 633,292 size 64x24; TextOff 'Back'
      on Click: ActivateScreen("Screen_3", 0)
   Button "Button_6" at 716,292 size 64x24; TextOff 'Next'
      on Click: ActivateScreen("Screen_5", 0)
   GraphicView "Template_Graphic view_1" at 736,255 size 28x26; Picture "NEW_HOME"
   GraphicView "Template_Graphic view_2" at 650,253 size 28x27; Picture "play"
   GraphicView "Template_Graphic view_3" at 721,296 size 20x17; Picture "next-track"
   GraphicView "Template_Graphic view_4" at 638,296 size 20x17; Picture "previous-track"
   Button "Button_3" at 707,246 size 80x42; TextOn 'LOGOUT'; TextOff 'Text'
      on Activate: function_f23ef4c9(); ActivateScreen("1_OVERVIEW_1", 0)
   Button "Button_1" at 623,245 size 80x42; TextOff 'Text'
      on Press: SetTag("มีการปุ่มกดยืนยัน", 1)
      on Release: SetTag("มีการปุ่มกดยืนยัน", 0)
      on Activate: "Storage"()
      on Click: "Conveyor"(); ActivateScreen("Status System", 0)
   TextField "Text field_49" at 734,229 size 32x14; Text 'HOME'
   TextField "Text field_50" at 625,229 size 95x16; Text 'Simmulation Conveyor'

